(* IEC 61131-3 sources: NachHouse_TST/OSCAT_BasicLib/OscatBasicLib_333a (part 5) *)

(* ---- Plc_Time.ST ---- *)
(* @PATH := '\/Engineering\/measurements' *)
FUNCTION T_PLC_MS : DWORD
(*
  T_PLC_MS reads the internal PLC timer and return the time, it has the advantage to be able to set a debug mode
  and speed up the counter to test the plc timer overrun which occurs every 50 days respectively 25 days at siemens S7
  this routine also allows to correct the behavior of s7 where the internal plc counter will not count all 32 bits.

  version 1.2 16. nov 2008
  programmer  hugo
  tested by oscat
*)
  VAR CONSTANT
    debug : BOOL := 0;
    N : INT := 0;
    offset : DWORD := 0;
  END_VAR
  VAR
  //  tx : TIME;
  END_VAR
  VAR_EXTERNAL
    AT %SL52 : DWORD;
  END_VAR
  VAR_TEMP
    temp : DWORD;
  END_VAR

  //???tx := TIME();
  T_PLC_MS := %SL52;
  (* hier muss die korrektur für step7 stattfinden
  plctime muss den vollen wertebereich von time ausnutzen:
  wenn bei step7 time -24tage bis plus 24 tage ist dann muss der timer auch beim überlauf auf -24tage springen
  und auf keinen fall auf 0 !!!!
  für siemens muss ein weiterer fb im main eingebunden werden der sicherstellt das alle 32 bits durchgezählt werden.
  es kann nur ein fb sein den er muss sich das oberste (32te) bit merken.
  oder etwa spring s7 bei überlauf auf -24 tage????? dann wäre keine korrektur nötig.
  *)
  IF debug THEN
    //???  T_PLC_MS := (SHL(T_PLC_MS,N) OR SHL(DWORD#1,N)-1) + OFFSET;
    temp := UDINT_TO_DWORD( DWORD_TO_UDINT( SHL(DWORD#1,INT_TO_UINT(N))) -1);
    temp := temp OR SHL(%SL52,INT_TO_UINT(N));
    T_PLC_MS := UDINT_TO_DWORD( DWORD_TO_UDINT(temp) + DWORD_TO_UDINT(OFFSET));
  END_IF;

(* revision history
  hm  14.9.2007 rev 1.0
    original version

  hm  12. nov 2007  rev 1.1
    added temporaray variable tx because some compilers could not handle time() as an argument

  hm  16. nov. 2008 rev 1.2
    initialized constants with 0 for compatibility reasons
*)
END_FUNCTION

(* @PATH := '\/Engineering\/measurements' *)
FUNCTION T_PLC_US : DWORD
(*
  T_PLC_US reads the internal PLC timer and return the time, it has the advantage to be able to set a debug mode
  and speed up the counter to test the plc timer overrun which occurs every 50 days respectively 25 days at siemens S7
  this routine also allows to correct the behavior of s7 where the internal plc counter will not count all 32 bits.

  version 1.2 16 nov 2008
  programmer  hugo
  tested by tobias
*)
  VAR CONSTANT
    debug : BOOL := 0;
    N : INT := 0;
    offset : DWORD := 0;
  END_VAR
  VAR
  //  tx : TIME;
  END_VAR
  VAR_EXTERNAL
    AT %SL52 : DWORD;
  END_VAR
  VAR_TEMP
    temp : DWORD;
    temp_T_PLC_US : DWORD;
  END_VAR

  //???tx := TIME();
  //???T_PLC_US := TIME_TO_DWORD(Tx)*1000;
  T_PLC_US := UDINT_TO_DWORD(DWORD_TO_UDINT(%SL52)*1000);
  (* hier muss die korrektur für step7 stattfinden
  plctime muss den vollen wertebereich von time ausnutzen:
  wenn bei step7 time -24tage bis plus 24 tage ist dann muss der timer auch beim überlauf auf -24tage springen
  und auf keinen fall auf 0 !!!!
  für siemens muss ein weiterer fb im main eingebunden werden der sicherstellt das alle 32 bits durchgezählt werden.
  es kann nur ein fb sein den er muss sich das oberste (32te) bit merken.
  oder etwa spring s7 bei überlauf auf -24 tage????? dann wäre keine korrektur nötig.
  *)
  IF debug THEN
    //???T_PLC_US := (SHL(T_PLC_US,N) OR SHL(DWORD#1,N)-1) + OFFSET;
    temp_T_PLC_US := UDINT_TO_DWORD(DWORD_TO_UDINT(%SL52)*1000);
    temp := UDINT_TO_DWORD( DWORD_TO_UDINT( SHL(DWORD#1,INT_TO_UINT(N))) -1);
    temp := temp OR SHL(temp_T_PLC_US,INT_TO_UINT(N));
    T_PLC_US := UDINT_TO_DWORD( DWORD_TO_UDINT(temp) + DWORD_TO_UDINT(OFFSET));
  END_IF;

(* revision history
  hm  14.9.2007 rev 1.0
    original version

  hm  12. nov 2007  rev 1.1
    added temporaray variable tx because some compilers could not handle time() as an argument

  hm  16. nov. 2008 rev 1.2
    initialized constants with 0 for compatibility reasons
*)
END_FUNCTION

(* @PATH := '\/String' *)
FUNCTION TO_UPPER : BYTE
(*
  to_upper converts a character from lowercase to uppercase

  version 1.3 16. jan. 2009
  programmer  hugo
  tested by   oscat
*)
  VAR_INPUT
    IN : BYTE;
  END_VAR

  IF (in > 96) AND (in < 123) THEN
     TO_UPPER := in AND 16#DF;
  ELSIF (in > 223) AND (in <> 247) AND (in <> 255) AND setup.EXTENDED_ASCII THEN
     TO_UPPER := in AND 16#DF;
  ELSE
     TO_UPPER := in;
  END_IF;

(* revision history
  hm  6. mar. 2008  rev 1.0
    original version

  hm  19. oct. 2008 rev 1.1
    changed setup constants

  ks  25. oct. 2008 rev 1.2
    optimized code

  hm 16. jan 2009 rev 1.3
    corrected an error in module
  *)
END_FUNCTION

(* ---- Sensors.ST ---- *)
(* @PATH := '\/Engineering\/sensor' *)
FUNCTION MULTI_IN : REAL
(*
  multi_in is a signal conditioning function which can be configured in 8 different ways.
  it is used to read multiple sensors for the same value and protect the user from broken sensors or invalid data from sensors.

  multi_in can be configured in different ways:
    mode = 0 means the the avg of the 3 inputs is used, this mode is the default mode.
    mode = 1 means in_1 is used.
    mode = 2 means in_2 is used.
    mode = 3 means in_3 is used.
    mode = 4 means default is used.
    mode = 5 means the lowest of the 3 external temperatures is used.
    mode = 6 means the higest externnal temperature is used.
    mode = 7 means the midlle input is used, if there are only two working, the lowest input is used.
    mode > 7 ,eans output is 0 at all times.
    in any config mode, an input higher then in_max or lower then in_min is ignored to prevent values from broken sensors or wires.
    if all inputs are higher then in_max or lower then in_min, a default value (default) is used.

  version 1.4 18. jul. 2009
  programmer  oscat
  tested by   oscat
*)
  VAR_INPUT
    in_1 : REAL;
    in_2 : REAL;
    in_3 : REAL;
    default : REAL;
    in_min : REAL;
    in_max : REAL;
    mode : BYTE;
  END_VAR
  VAR
    count: INT;
    F1: BOOL;
    F2: BOOL;
    F3: BOOL;
  END_VAR

  F1 :=  in_1 > in_min AND in_1 < in_max;
  F2 :=  in_2 > in_min AND in_2 < in_max;
  F3 :=  in_3 > in_min AND in_3 < in_max;

  CASE BYTE_TO_USINT(mode) OF
  0:  count := 0;
    IF F1 THEN
      count := count + 1;
      MULTI_IN := in_1;
    ELSE
      MULTI_IN := 0.0;
    END_IF;
    IF F2 THEN
      count := count + 1;
      MULTI_IN := MULTI_IN + in_2;
    END_IF;
    IF F3 THEN
      count := count + 1;
      MULTI_IN := MULTI_IN + in_3;
    END_IF;
    MULTI_IN := SEL(count = 0, MULTI_IN / INT_TO_REAL(count), default);

  1:  MULTI_IN := SEL(F1, default, IN_1);

  2:  MULTI_IN := SEL(F2, default, IN_2);

  3:  MULTI_IN := SEL(F3, default, IN_3);

  4:  MULTI_IN := default;

  5:  MULTI_IN := SEL(F1, in_max, IN_1);
    IF F2 AND in_2 < MULTI_IN THEN MULTI_IN := in_2; END_IF;
    IF F3 AND in_3 < MULTI_IN THEN MULTI_IN := in_3; END_IF;
    IF MULTI_IN = in_max THEN MULTI_IN := default; END_IF;

  6:  MULTI_IN := SEL(F1, in_min, IN_1);
    IF F2 AND in_2 > MULTI_IN THEN MULTI_IN := in_2; END_IF;
    IF F3 AND in_3 > MULTI_IN THEN MULTI_IN := in_3; END_IF;
    IF MULTI_IN = in_min THEN MULTI_IN := default; END_IF;

  7:  IF F1 AND F2 AND F3 THEN MULTI_IN := MID3(in_1, in_2, in_3);
    ELSIF F1 AND F2 THEN MULTI_IN := MIN(in_1, in_2);
    ELSIF F1 AND F3 THEN MULTI_IN := MIN(in_1, in_3);
    ELSIF F2 AND F3 THEN MULTI_IN := MIN(in_2, in_3);
    ELSIF F1 THEN MULTI_IN := in_1;
    ELSIF F2 THEN MULTI_IN := in_2;
    ELSIF F3 THEN MULTI_IN := in_3;
    ELSE MULTI_IN := default;
    END_IF;
  ELSE
    MULTI_IN := 0.0;
  END_CASE;

(*
  hm 1.1.2007   rev 1.1
    changed midr to mid3 function

  hm  14. 10. 2008  rev 1.2
    corrected an error for in_3 overrange detection
    improved performance

  hm  11. mar. 2009 rev 1.3
    changed real constants to use dot syntax

  hm  18. jul. 2009 rev 1.4
    improved performance
*)
END_FUNCTION

(* @PATH := '\/Engineering\/sensor' *)
FUNCTION RES_NI : REAL
(*
  this function returs the resistance for a nickel sensor for a temperature range from -60..+180 °C

  version 1.2 2 dec 2007
  programmer  hugo
  tested by   tobias
*)
  VAR_INPUT
    T : REAL;
    R0 : REAL;
  END_VAR
  VAR CONSTANT
    A : REAL := 0.5485;
    B : REAL := 0.665E-3;
    C : REAL := 2.805E-9;
  END_VAR
  VAR
    T2: REAL;
  END_VAR

  T2 := T * T;
  RES_NI := R0 + A * T + B * T2 + C * T2 * T2;

(* revision history
  hm  4.8.2006    rev 1.0
    original version

  hm  13.9.2007   rev 1.1
    changed coding for better performance

  hm  2. dec. 2007  rev 1.2
    changed code for better performance
*)
(*
 Auszug aus DIN 43760 für Ni100

°C    R   °C    R   °C  R   °C    R   °C    R

-60   69,5  -10   94,6  40  123,0   90    154,9   140   190,9
-55   71,9  -5    97,3  45  126,0   95    158,3   145   194,8
-50   74,3  0     100,0   50  129,1   100   161,8   150   198,7
-45   76,7  5     102,8   55  132,2   105   165,3   155   202,6
-40   79,1  10    105,6   60  135,3   110   168,8   160   206,6
-35   81,6  15    108,4   65  138,5   115   172,4   165   210,7
-30   84,2  20    111,2   70  141,7   120   176,0   170   214,8
-25   86,7  25    114,1   75  145,0   125   179,6   175   219,0
-20   89,3  30    117,1   80  148,3   130   183,3   180   223,2
-15   91,9  35    120,0   85  151,6   135   187,1
*)
END_FUNCTION

(* @PATH := '\/Engineering\/sensor' *)
FUNCTION RES_NTC : REAL
(*
  this function returs the resistance for a NTC sensor for a given temperature in °C.
  RN is the resistance at 25 °C and B is a constant for the given sensor.

  version 1.1 11. mar. 2009
  programmer  hugo
  tested by   tobias
*)
  VAR_INPUT
    T : REAL;
    RN : REAL;
    B : REAL;
  END_VAR

  RES_NTC := RN * EXP(B * (1.0 / (T+273.15) - 0.00335401643468053));

(* revision history
  hm 30. dec. 2008  rev 1.0
    original version

  hm  11. mar. 2009 rev 1.1
    changed real constants to use dot syntax
*)
END_FUNCTION

(* @PATH := '\/Engineering\/sensor' *)
FUNCTION RES_PT : REAL
(*
  this function returs the resistance for a platinum sensor for a temperature range from -200..+850 °C

  version 1.3 11. mar. 2009
  programmer  hugo
  tested by   oscat
*)
  VAR_INPUT
    T : REAL;
    R0 : REAL;
  END_VAR
  VAR CONSTANT
    A : REAL := 3.90802E-3 ;
    B : REAL := -5.802E-7;
    C : REAL := -4.27350E-12;
  END_VAR
  VAR
    T2: REAL;
  END_VAR

  T2 := T * T;

  IF T >= 0.0 THEN
    RES_PT := R0 * ( 1.0 + A * T + B * T2);
  ELSE
    RES_PT := R0 * ( 1.0 + A * T + B * T2 + C * (T - 100.0) * T2 * T);
  END_IF;

(* revision history
  hm  4. aug. 2006  rev 1.1
    original version

  hm  2. dec 2007 rev 1.2
    changed code for better performance

  hm  11. mar. 2009 rev 1.3
    changed real constants to use dot syntax
*)
(*
 Auszug aus DIN 43760 für Pt100

°C    R   °C    R   °C  R     °C    R     °C    R     °C    R

-200  18,49   -100  60,25   0   100,00  100   138,50  200   175,84  300   212,02
-195  20,65   -95   62,28   5   101,95  105   140,39  205   177,68  305   213,80
-190  22,80   -90   64,30   10  103,90  110   142,29  210   179,51  310   215,57
-185  24,94   -85   66,31   15  105,85  115   144,17  215   181,34  315   217,35
-180  27,08   -80   68,33   20  107,79  120   146,06  220   183,17  320   219,12
-175  29,20   -75   70,33   25  109,73  125   147,94  225   184,99  325   220,88
-170  31,32   -70   72,33   30  111,67  130   149,82  230   186,82  330   222,65
-165  33,43   -65   74,33   35  113,61  135   151,70  235   188,63  335   224,41
-160  35,33   -60   76,33   40  115,54  140   153,58  240   190,45  340   226,17
-155  37,63   -55   78,32   45  117,47  145   155,45  245   192,26  345   227,92
-150  39,71   -50   80,31   50  119,40  150   157,31  250   194,07  350   229,67
-145  41,79   -45   82,29   55  121,32  155   159,18  255   195,88  355   231,42
-140  43,87   -40   84,27   60  123,24  160   161,04  260   197,69  360   233,17
-135  45,94   -35   86,25   65  125,16  165   162,90  265   199,49  365   234,91
-130  48,00   -30   88,22   70  127,07  170   164,76  270   201,29  370   236,65
-125  50,06   -25   90,19   75  128,98  175   166,61  275   203,08  375   238,39
-120  52,11   -20   92,16   80  130,89  180   168,46  280   204,88  380   240,13
-115  54,15   -15   94,12   85  132,80  185   170,31  285   206,67  385   241,86
-110  56,19   -10   96,09   90  134,70  190   172,16  290   208,45  390   243,59
-105  58,22   -5    98,04   95  136,60  195   174,00  295   210,24  395   245,31
*)
END_FUNCTION

(* @PATH := '\/Engineering\/sensor' *)
FUNCTION RES_SI : REAL
(*
  this function returs the resistance for a silicon sensor for a temperature range from -50..+150 °C
  for example KTY10 normaly Rs at 25 °C

  version 1.2 11. mar. 2009
  programmer  hugo
  tested by   tobias
*)
  VAR_INPUT
    T : REAL;
    RS : REAL;
    TS : REAL;
  END_VAR
  VAR CONSTANT
    A : REAL := 7.64E-3;
    B : REAL := 1.66E-5;
  END_VAR
  VAR
    TX: REAL;
  END_VAR

  TX := T - TS;
  RES_SI := RS * ( 1.0 + A * TX + B * TX * TX);

(* revision history
  hm  4. aug 2006 rev 1.0
    original version

  hm  2. dec 2007 rev 1.1
    changed code for better performance

  hm  11. mar. 2009 rev 1.2
    changed real constants to use dot syntax
*)
END_FUNCTION

(* @PATH := '\/Engineering\/sensor' *)
FUNCTION SENSOR_INT : REAL
(*
  this function calculates the real resistance of a sensor RX given a parasitic resistor in parallel to the sensor and an additional serial resistor.
  for example a parasitic parallel resistor for a PT100 can be ignored but a series resistor is the cable to the sensor.
  for a humidity sensor, the parallel resistor is more dramatic and needs to be considered.
  the function allows to consider a parallel and serial resistor at the same time.
  with this function and known parasitic serial and parallel resistors the true resistance of the sensor can be calculated.

  version 1.3 11. mar. 2009
  programmer  hugo
  tested by   tobias
*)
  VAR_INPUT
    Voltage : REAL;
    Current : REAL;
    RP : REAL;
    RS : REAL;
  END_VAR
  VAR
    RG: REAL;
  END_VAR

  IF current <> 0.0 THEN
    RG := voltage / current;
    SENSOR_INT := RP * ( RG - RS) / ( RP + RS - RG);
  END_IF;

(* revisaion history
  hm 20.1.2007    rev 1.1
    deleted input R0 which was not needed.

  hm  2. dec 2007 rev 1.2
    corrected an error in formula and improoved speed

  hm  11. mar. 2009 rev 1.3
    changed real constants to use dot syntax
*)
END_FUNCTION

(* @PATH := '\/Engineering\/sensor' *)
FUNCTION TEMP_NI : REAL
(*
  this function returns the temperature for a nickel sensor in a range from -60..+180 °C

  version 1.5 10. mar. 2009
  programmer  hugo
  tested by   tobias
*)
  VAR_INPUT
    Res : REAL;
    R0 : REAL;
  END_VAR

  TEMP_NI := (SQRT(0.30085225 - 2.66E-3 * (R0 - Res)) - 0.5485) * 751.8796992;

(* revision history
  hm 24.1.2007    rev 1.1
    deleted unused variable A, B, C

  hm 10.9.2007    rev 1.2
    changed accuracy to 0.02 degrees to improove performace

  hm 17. 12 2007  rev 1.3
    improovements for better performance and higher accuracy

  hm  6. jan 2008 rev 1.4
    further performance improvement

  hm  10. mar. 2009 rev 1.5
    removed nested comments
*)
END_FUNCTION

(* @PATH := '\/Engineering\/sensor' *)
FUNCTION TEMP_NTC : REAL
(*
  this function returs the temperature for a NTC sensor for a range from 0..85 °C.
  RN is the resistance at 25 °C and B is a constant for the given sensor.

  version 1.1 11. mar. 2009
  programmer  hugo
  tested by   tobias
*)
  VAR_INPUT
    RES : REAL;
    RN : REAL;
    B : REAL;
  END_VAR

  IF res > 0.0 THEN
    TEMP_NTC := B * 298.15 / (B + LN(RES / RN) * 298.15) -273.15;
  END_IF;

(* revision history
  hm 30. dec. 2008  rev 1.0
    original version

  hm  11. mar. 2009 rev 1.1
    changed real constants to use dot syntax
*)
END_FUNCTION

(* @PATH := '\/Engineering\/sensor' *)
FUNCTION TEMP_PT : REAL
(*
  this function returs the temperature for a platinum sensor for a range from -200..+850 °C

  version 1.7 11. mar. 2009
  programmer  hugo
  tested by   oscat
*)
  VAR_INPUT
    Res : REAL;
    R0 : REAL;
  END_VAR
  VAR CONSTANT
    A : REAL := 3.9083E-3 ;
    B : REAL := -5.775E-7;
    accuracy : REAL := 0.01;
  END_VAR
  VAR
    step: REAL := 50.0;
    X: REAL;
    Y: REAL;
    t1: REAL;
    pt : PTR_TO UDINT; //DWORD;
  END_VAR
  VAR_TEMP
    tmp : REAL;
  END_VAR

  X := A * R0;
  Y := B * R0;
  IF Res >= R0 THEN
    t1 := X * X - 4.0 * Y * (R0 - Res);
    IF t1 < 0.0 THEN
      tmp := 10000.0;
    ELSE
      tmp := (-X + SQRT(t1)) / (2.0 * Y);
    END_IF;
  ELSE
    pt := ADR(step);
    (* since the formula cannot be solved this is a successive approximation *)
    tmp := -100.0;
    WHILE step > accuracy DO
      (* test if result greater or less *)
      IF RES_PT(tmp, R0) < res THEN tmp := tmp + step; ELSE tmp := tmp - step; END_IF;
      pt^ := pt^ - 8388608;  (* this is a super fast divide by 2 method for non floating point CPUs *)
      (* the alternative code: step := step * 0.5; *)
    END_WHILE;
  END_IF;
  TEMP_PT := tmp;

(* revision history
  rev 1.1 hm 24.1.2007
    deleted unused variable C

  rev 1.2 hm 10.9.2007
    reduced accuracy to 0.02 to shorten execution time

  rev 1.3 hm  2. dec 2007
    changed code for better performance

  rev 1.4 hm  23. dec 2007
    avoid a negative square root if input values are wrong

  rev 1.5 hm  5. jan 2008
    replaced / 2 with * 0.5 for better performance

  hm  31. oct. 2008 rev 1.6
    improved performance

  hm  11. mar. 2009 rev 1.7
    changed real constants to use dot syntax
*)
END_FUNCTION

(* @PATH := '\/Engineering\/sensor' *)
FUNCTION TEMP_SI : REAL
(*
  this function returs the temperature for a silicon sensor for a range from -60..+180 °C
  for example KTY10 RS at TS normally 25 °C

  version 1.5 10. mar. 2009
  programmer  hugo
  tested by   tobias
*)
  VAR_INPUT
    Res : REAL;
    RS : REAL;
    TS : REAL;
  END_VAR

  TEMP_SI := (-7.64E-3 + SQRT(Res / RS * 6.64E-5 - 0.803E-5)) * 30120.48193 + TS;

(* revision history
  hm 24.1.2007    rev 1.1
    the function would only work for TS = 25, now it works for other values of ts.

  hm 10.9.2007    rev 1.2
    changed the function to use successive approcimation to avoid an error generated by a sqrt from a negative result.
    changed accuracy to 0.02 degrees to shorten execution time

  hm 17. 12 2007  rev 1.3
    improovements for better performance

  hm  6. jan 2008 rev 1.4
    further performance improvement

  hm  10. mar. 2009 rev 1.5
    removed nested comments
*)
END_FUNCTION

(* ---- String.ST ---- *)
(* @NESTEDCOMMENTS := 'Yes' *)
(* @PATH := '\/String' *)
(* @OBJECTFLAGS := '0, 8' *)
(* @SYMFILEFLAGS := '2048' *)
FUNCTION TO_UPPER : BYTE
(*
  to_upper converts a character from lowercase to uppercase

  version 1.3 16. jan. 2009
  programmer  hugo
  tested by   oscat
*)
  VAR_INPUT
    IN : BYTE;
  END_VAR

  (* @END_DECLARATION := '0' *)
  IF BYTE_TO_USINT(in) > 96 AND BYTE_TO_USINT(in) < 123 THEN
     TO_UPPER := in AND 16#DF;
  ELSIF BYTE_TO_USINT(in) > 223 AND BYTE_TO_USINT(in) <> 247 AND BYTE_TO_USINT(in) <> 255 AND setup.EXTENDED_ASCII THEN
     TO_UPPER := in AND 16#DF;
  ELSE
     TO_UPPER := in;
  END_IF;

  (* revision history
  hm  6. mar. 2008  rev 1.0
    original version

  hm  19. oct. 2008 rev 1.1
    changed setup constants

  ks  25. oct. 2008 rev 1.2
    optimized code

  hm 16. jan 2009 rev 1.3
    corrected an error in module

  *)
END_FUNCTION

(* ---- Vector_Mathematics.ST ---- *)
(* @PATH := '\/Mathematical\/Vektormathematik' *)
FUNCTION V3_ABS : REAL
(*
  this function calculates the length of a vectors in a 3 dimensional space

  version 1.0 11 dec 2007
  programmer  hugo
  tested by   tobias
*)
  VAR_INPUT
    A : Vector_3;
  END_VAR

  V3_ABS := SQRT(A.X * A.X + A.Y * A.Y + A.Z * A.Z);

(* revision history
  hm  11 dec 2007 rev 1.0
      original version
*)
END_FUNCTION

(* @PATH := '\/Mathematical\/Vektormathematik' *)
FUNCTION V3_ADD : vector_3
(*
  this function adds two vectors in a 3 dimensional space

  version 1.0 11 dec 2007
  programmer  hugo
  tested by   tobias
*)
  VAR_INPUT
    A : Vector_3;
    B : Vector_3;
  END_VAR

  V3_ADD.X := A.X + B.X;
  V3_ADD.Y := A.Y + B.Y;
  V3_ADD.Z := A.Z + B.Z;

(* revision history
  hm    11 dec 2007 rev 1.0
        original version
*)
END_FUNCTION

(* @PATH := '\/Mathematical\/Vektormathematik' *)
FUNCTION V3_DPRO : REAL
(*
  this function calculates the dot product of two vectors in 3 dimensional space

  version 1.0 11 dec 2007
  programmer  hugo
  tested by   tobias
*)
  VAR_INPUT
    A : Vector_3;
    B : Vector_3;
  END_VAR

  V3_DPRO := A.X * B.X + A.Y * B.Y + A.Z * B.Z;

(* revision history
  hm  11 dec 2007 rev 1.0
      original version
*)
END_FUNCTION

(* @PATH := '\/Mathematical\/Vektormathematik' *)
FUNCTION V3_ANG : REAL
(*
  this function calculates the angle between two vectors in a 3 dimensional space

  version 1.1 10. mar. 2009
  programmer  hugo
  tested by   tobias
*)
  VAR_INPUT
    A : Vector_3;
    B : Vector_3;
  END_VAR
  VAR
    d : REAL;
  END_VAR

  d := V3_ABS(A) * V3_ABS(B);
  IF d > 0.0 THEN
    V3_ANG := ACOS(LIMIT(-1.0, V3_DPRO(A, B) / d,1.0));
  END_IF;

(* revision history
  hm  11. dec. 2007 rev 1.0
    original version

  hm  10. mar. 2009 rev 1.1
    changed syntax of real constants to 0.0
*)
END_FUNCTION

(* @PATH := '\/Mathematical\/Vektormathematik' *)
FUNCTION V3_SMUL : vector_3
(*
  this function multiplies a vectors in a 3 dimensional space with a skalar M

  version 1.0 11 dec 2007
  programmer  hugo
  tested by   tobias
*)
  VAR_INPUT
    A : Vector_3;
    M : REAL;
  END_VAR

  V3_SMUL.X := A.X * M;
  V3_SMUL.Y := A.Y * M;
  V3_SMUL.Z := A.Z * M;

(* revision history
  hm    11 dec 2007 rev 1.0
        original version
*)
END_FUNCTION

(* @PATH := '\/Mathematical\/Vektormathematik' *)
FUNCTION V3_NORM : vector_3
(*
  this function generates a vectors with absolute length 1 from a vector A in a 3 dimensional space

  version 1.1 10. mar. 2009
  programmer  hugo
  tested by   tobias
*)
  VAR_INPUT
    A : Vector_3;
  END_VAR
  VAR
    la: REAL;
  END_VAR

  la := V3_ABS(A);
  IF la > 0.0 THEN
    V3_NORM := V3_SMUL(A, 1.0 / la);
  END_IF;

(* revision history
  hm  11 dec 2007 rev 1.0
    original version

  hm  10. mar. 2009 rev 1.1
    changed syntax of real constants to 0.0
*)
END_FUNCTION

(* @PATH := '\/Mathematical\/Vektormathematik' *)
FUNCTION V3_NUL : BOOL
(*
  this function checks if a vectors in a null Vector

  version 1.1 10. mar. 2009
  programmer  hugo
  tested by   tobias
*)
  VAR_INPUT
    A : Vector_3;
  END_VAR

  V3_NUL := A.X = 0.0 AND A.Y = 0.0 AND A.Z = 0.0;

(* revision history
  hm  12 dec 2007 rev 1.0
    original version

  hm  10. mar. 2009 rev 1.1
    changed syntax of real constants to 0.0
*)
END_FUNCTION

(* @PATH := '\/Mathematical\/Vektormathematik' *)
FUNCTION V3_XPRO : vector_3
(*
  this function adds two vectors in a 3 dimensional space

  version 1.0 11 dec 2007
  programmer  hugo
  tested by   tobias
*)
  VAR_INPUT
    A : Vector_3;
    B : Vector_3;
  END_VAR

  V3_XPRO.X := A.Y * B.Z - A.Z * B.Y;
  V3_XPRO.Y := A.Z * B.X - A.X * B.Z;
  V3_XPRO.Z := A.X * B.Y - A.Y * B.X;

(* revision history
  hm    11 dec 2007 rev 1.0
    original version
*)
END_FUNCTION

(* @PATH := '\/Mathematical\/Vektormathematik' *)
FUNCTION V3_PAR : BOOL
(*
  this function checks if two vectors in a 3 dimensional space are parallel.
  which means the two vectors have the same direction

  version 1.1 10. mar. 2009
  programmer  hugo
  tested by   tobias
*)
  VAR_INPUT
    A : Vector_3;
    B : Vector_3;
  END_VAR

  V3_PAR := V3_ABS(V3_XPRO(A, B)) = 0.0;

(* revision history
  hm  11 dec 2007 rev 1.0
    original version

  hm  10. mar. 2009 rev 1.1
    changed syntax of real constants to 0.0
*)
END_FUNCTION

(* @PATH := '\/Mathematical\/Vektormathematik' *)
FUNCTION V3_REV : vector_3
(*
  this function reverses a vector in a 3 dimensional space

  version 1.0 11 dec 2007
  programmer  hugo
  tested by   tobias
*)
  VAR_INPUT
    A : Vector_3;
  END_VAR

  V3_REV.X := -A.X;
  V3_REV.Y := -A.Y;
  V3_REV.Z := -A.Z;

(* revision history
  hm    11 dec 2007 rev 1.0
        original version
*)
END_FUNCTION

(* @PATH := '\/Mathematical\/Vektormathematik' *)
FUNCTION V3_SUB : vector_3
(*
  this function subtracts two vectors in a 3 dimensional space
  V3_SUB = A - B

  version 1.0 11 dec 2007
  programmer  hugo
  tested by   tobias
*)
  VAR_INPUT
    A : Vector_3;
    B : Vector_3;
  END_VAR

  V3_SUB.X := A.X - B.X;
  V3_SUB.Y := A.Y - B.Y;
  V3_SUB.Z := A.Z - B.Z;

(* revision history
  hm    11 dec 2007 rev 1.0
    original version
*)
END_FUNCTION

(* @PATH := '\/Mathematical\/Vektormathematik' *)
FUNCTION V3_XANG : REAL
(*
  this function calculates the angle between the X-axis and a vectors in a 3 dimensional space

  version 1.1 10. mar. 2009
  programmer  hugo
  tested by   tobias
*)
  VAR_INPUT
    A : Vector_3;
  END_VAR
  VAR
    la: REAL;
  END_VAR

  la := V3_ABS(a);
  IF la > 0.0 THEN
    V3_XANG := ACOS(A.X / la);
  END_IF;

(* revision history
  hm  11 dec 2007 rev 1.0
    original version

  hm  10. mar. 2009 rev 1.1
    changed syntax of real constants to 0.0
*)
END_FUNCTION

(* @PATH := '\/Mathematical\/Vektormathematik' *)
FUNCTION V3_YANG : REAL
(*
  this function calculates the angle between the Y-axis and a vectors in a 3 dimensional space

  version 1.1 10. mar. 2009
  programmer  hugo
  tested by   tobias
*)
  VAR_INPUT
    A : Vector_3;
  END_VAR
  VAR
    la: REAL;
  END_VAR

  la := V3_ABS(a);
  IF la > 0.0 THEN
    V3_YANG := ACOS(A.Y / la);
  END_IF;

(* revision history
  hm  11 dec 2007 rev 1.0
    original version

  hm  10. mar. 2009 rev 1.1
    changed syntax of real constants to 0.0
*)
END_FUNCTION

(* @PATH := '\/Mathematical\/Vektormathematik' *)
FUNCTION V3_ZANG : REAL
(*
  this function calculates the angle between the Z-axis and a vectors in a 3 dimensional space

  version 1.1 10. mar. 2009
  programmer  hugo
  tested by   tobias
*)
  VAR_INPUT
    A : Vector_3;
  END_VAR
  VAR
    la: REAL;
  END_VAR

  la := V3_ABS(a);
  IF la > 0.0 THEN
    V3_ZANG := ACOS(A.Z / la);
  END_IF;

(* revision history
  hm  11 dec 2007 rev 1.0
    original version

  hm  10. mar. 2009 rev 1.1
    changed syntax of real constants to 0.0
*)
END_FUNCTION

(* ---- Arithmetic_Functions.ST ---- *)
TYPE
  OSCAT_BASIC_ARRAY1_20x0_1_OF_REAL : ARRAY[1..20, 0..1] OF REAL;
END_TYPE

(* @PATH := '\/Mathematical\/functions' *)
FUNCTION F_LIN : REAL
(*
  this function calculates the linear equation f_lin = a*x + b

  version 1.0 1 sep 2006
  programmer  hugo
  tested by   tobias
*)
  VAR_INPUT
    X : REAL;
    A : REAL;
    B : REAL;
  END_VAR

  F_lin := A * X + B;
END_FUNCTION

(* @PATH := '\/Mathematical\/functions' *)
FUNCTION F_LIN2 : REAL
(*
  this function calculates the linear equation f_lin = a*x + b given by two points x1/y1 and x2/y2.

  version 1.0 1 jan 2007
  programmer  hugo
  tested by   tobias
*)
  VAR_INPUT
    X : REAL;
    X1: REAL;
    Y1 : REAL;
    X2 : REAL;
    Y2 : REAL;
  END_VAR

  F_LIN2 := (Y2 - Y1) / (X2 - X1) * (X - X1) + Y1;

(* revision history
  hm  1. jan. 2007  rev 1.0
    original release

  hm  17. dec. 2008 rev 1.1
    optimized formula
*)
END_FUNCTION

(* @PATH := '\/Mathematical\/functions' *)
FUNCTION F_POLY : REAL
(*
  this function calculates the polynom C[0] + C[1]*X^1 + C[2]*X^2 * C[3]*X^3 + C[4]*X^4 + C[5]*X^5 + C[6]*X^6 + C[7]*X^7

  version 1.1 18. mar. 2011
  programmer  hugo
  tested by   tobias
*)
  VAR_INPUT
    X : REAL;
    C : ARRAY[0..7] OF REAL;
  END_VAR

  F_POLY := ((((((( c[7] * x + c[6] ) * x + c[5] ) * x + c[4] ) * x + c[3] ) * x + c[2] ) * x + c[1] ) * x + c[0] ) ;

(* revision history
  hm    20. may. 2008   rev 1.0
    original version

  hm  18. mar. 2011 rev 1.1
    improved performance
*)
END_FUNCTION

(* @PATH := '\/Mathematical\/functions' *)
FUNCTION F_POWER : REAL
(*
  this function calculates the power equation f_power = a*x^n

  version 1.0 1 sep 2006
  programmer  hugo
  tested by   tobias
*)
  VAR_INPUT
    a : REAL;
    x : REAL;
    n : REAL;
  END_VAR

  F_POWER := a * EXPT(X, N);
END_FUNCTION

(* @PATH := '\/Mathematical\/functions' *)
FUNCTION F_QUAD : REAL
(*
  this function calculates the quadratic equation f_lin = a*x + b

  version 1.1 18. Mar. 2011
  programmer  hugo
  tested by   tobias
*)
  VAR_INPUT
    X : REAL;
    A : REAL;
    B : REAL;
    C : REAL;
  END_VAR

  F_QUAD :=  (A * X + B) * X + C;

(* revision history
  hm  1. sep. 2006  rev 1.0
    original version

  hm  18. mar. 2001 rev 1.1
    improved performance
*)
END_FUNCTION

(* @PATH := '\/Mathematical\/functions' *)
FUNCTION FRMP_B : BYTE
(*
  this function calculates a ramp and limits the output to 0 .. 255 without overflow problems

  version 1.0   17. feb. 2011
  programmer  hugo
  tested by   oscat
*)
  VAR_INPUT
    START : BYTE;
    DIR : BOOL;
    TD : TIME;
    TR : TIME;
  END_VAR
  VAR
    tmpw : DWORD;
    tmpb : BYTE;
  END_VAR

  IF TD < TR THEN
    //???FRMP_B := MIN(DWORD_TO_BYTE(SHL(TIME_TO_DWORD(TD), 8) / TIME_TO_DWORD(TR)), SEL(DIR, START, BYTE#255 - START));
    tmpw := SHL(TIME_TO_DWORD(TD), 8);
    tmpw := UDINT_TO_DWORD( DWORD_TO_UDINT(tmpw) /  TIME_TO_UDINT(TR));
    tmpb := MIN( DWORD_TO_BYTE(tmpw), SEL( DIR, START, USINT_TO_BYTE(USINT#255 - BYTE_TO_USINT(START))));
    IF DIR THEN
      FRMP_B := USINT_TO_BYTE( BYTE_TO_USINT(START) + BYTE_TO_USINT(tmpb));
    ELSE
      FRMP_B := USINT_TO_BYTE( BYTE_TO_USINT(START) - BYTE_TO_USINT(tmpb));
    END_IF;
  ELSE
    FRMP_B := SEL(DIR, 0, 255);
  END_IF;

(* revision history
  17. feb. 2011 rev 1.0
    new module
*)
END_FUNCTION

(* @PATH := '\/Mathematical\/functions' *)
FUNCTION_BLOCK FT_AVG
(*
  this function calculates the moving average over n samples from a sequential input
  the input values are shifted into an N deep buffer and the avg of this buffer is diplayed at anytime on the output.
  a rst will load the buffer with the current in value..

  version 1.5 10. mar. 2009
  programmer  hugo
  tested by   oscat
*)
  VAR_INPUT
    IN : REAL;
    E : BOOL := TRUE;
    N : INT := 32;
    RST : BOOL;
  END_VAR
  VAR_OUTPUT
    AVG : REAL;
  END_VAR
  VAR
    buff : DELAY;
    i: INT;
    init : BOOL;
  END_VAR

  (* limit n to a max of 32 because delay can do max 32 cycles *)
  buff.N := LIMIT(0, N, 32);

  IF NOT init OR rst THEN
    FOR i := 1 TO N DO
      buff(in := in);
    END_FOR;
    avg := in;
    init := TRUE;
  ELSIF E THEN
    buff(in := in);
    avg := avg + (in - buff.out ) / INT_TO_REAL(N);
  END_IF;

(* revision history
  hm  7. jan. 2007  rev 1.1
    chaged rst logic to load the buffer with the actual input value instead of 0.
    added en input to allow better control of signal flow
    added init to load the buffer with in at startup to avoid rampup at beginning.
    deleted unused variable cnt.

  hm  14. jun. 2008 rev 1.2
    set default for input en = TRUE and N = 32

  hm  10. oct. 2008 rev 1.3
    improved performance

  hm  18. oct. 2008 rev 1.4
    changed input en to e for compatibility reasons

  hm  10. mar. 2009 rev 1.5
    added type conversion for compatibility reasons
*)
END_FUNCTION_BLOCK

(* @PATH := '\/Mathematical\/functions' *)
FUNCTION_BLOCK FT_MIN_MAX
(*
  this function block stores the min and max value of an input signal.
  when rst is true the mn and mx outputs are set to the in value.
  when a rst is never active the function autoresets to the in value at startup.
  since the input might not be present at first cycle the mn and mx are set during second cycle.

  version 1.0 1 sep 2006
  programmer  hugo
  tested by   tobias
*)
  VAR_INPUT
    in : REAL;
    rst : BOOL;
  END_VAR
  VAR_OUTPUT
    mx : REAL;
    mn : REAL;
  END_VAR
  VAR
    init: BOOL;
  END_VAR

  IF rst OR NOT init THEN
    mn := in;
    mx := in;
    init := TRUE;
  ELSIF in < mn THEN mn := in;
  ELSIF in > mx THEN mx := in;
  END_IF;
END_FUNCTION_BLOCK

(* @PATH := '\/Mathematical\/functions' *)
FUNCTION_BLOCK FT_RMP
(*
  this ramp function follows an input signal with a linear ramp up or down, the up or down speed can be set with KF and KR.
  a K factor of 1 means 1 unit per second on the output. K factors can only be positive and not negative.
  a busy output signals the ramp is running or busy false means the in value is present on the output.
  a rmp input false means the output follows the input dierctly while a rmp = true means the output follows the input with a ramp.
  a updn output signal the directon of the ramp (up or down).

  version 1.4 25 jan 2008
  programmer  oscat
  tested by   oscat
*)
  VAR_INPUT
    Rmp : BOOL := TRUE;
    in : REAL;
    KR : REAL;
    KF : REAL;
  END_VAR
  VAR_OUTPUT
    out : REAL;
    busy : BOOL;
    UD : BOOL;
  END_VAR
  VAR
    tx: TIME;
    last: TIME;
    init: BOOL;
  END_VAR

  (* read system time *)
  tx := DWORD_TO_TIME(T_PLC_MS()) - last;

  IF NOT init THEN
    init := TRUE;
    last := tx;
    tx := t#0s;
    out := in;
  END_IF;
  IF NOT rmp THEN
    out := in;
    busy := FALSE;
  ELSIF out > in THEN
    (* ramp down *)
    out := out - TIME_TO_REAL(tx) * 0.001 * KF;
    out := MAX(in, out);
  ELSIF out < in THEN
    (* ramp up *)
    out := out + TIME_TO_REAL(tx) * 0.001 * KR;
    out := MIN(in, out);
  END_IF;

  (* set busy and dir flags *)
  IF out < in THEN
    busy := TRUE;
    ud := TRUE;
  ELSIF out > in THEN
    busy := TRUE;
    ud := FALSE;
  ELSE
    busy := FALSE;
  END_IF;
  last := last + tx;

(* revision history:
  hm 8.10.2006      rev 1.1
    added ud output

  hm 12. feb 2007   rev 1.2
    added init variable and corrected a possible startup problem

  hm  17. sep 2007  rev 1.3
    replaced time() with t_plc_ms() for compatibility reasons

  hm  25. jan 2008  rev 1.4
    performance improvements
    allow KR and KF to be 0
*)
END_FUNCTION_BLOCK

(* @PATH := '\/Mathematical\/functions' *)
FUNCTION LINEAR_INT : REAL
(*
  LINEAR_INT calculates an output based on a linear interpolation of up to 20 coordinates given in an array
  the input coordinates have to start at the lowest array position and must be sorted ba ascending X values.

  version 1.1 27 dec 2007
  programmer  oscat
  tested by   oscat
*)
  VAR_INPUT
    X : REAL;
    XY : OSCAT_BASIC_ARRAY1_20x0_1_OF_REAL; //ARRAY[1..20, 0..1] OF REAL;
    Pts : INT;
  END_VAR
  VAR
    i : INT;
  END_VAR

  (*make sure n is bound within the array size *)
  pts := MIN(pts,20);

  (* calculate the linear segement interpolation *)
  i := 2;
  (* search for segment and calculate output
    below and above the defined segments we interpolate the last segment *)
  WHILE (i < pts) AND (XY[i,0] < X) DO
    i := i + 1;
  END_WHILE;

  (* calculate the output value on the corresponding segment coordinates *)
  LINEAR_INT := ((XY[i,1] - XY[i-1,1]) * X - XY[i,1] * XY[i-1,0] + XY[i-1,1] * XY[i,0]) / (XY[i,0] - XY[i-1,0]);

(* revision history
  hm  7. oct 2007   rev 1.0
    original version

  hm  27 dec 2007   rev 1.1
    changed code for better performance
*)
END_FUNCTION

(* @PATH := '\/Mathematical\/functions' *)
FUNCTION POLYNOM_INT : REAL
(*
  POLYNOM_INT calculates an output based on a Polynom interpolation of up to 5 coordinates given in an array
  the indut coordinates have to start at the lowest array position and must be sorted ba ascending X values.

  version 1.3 10. mar. 2009
  programmer  oscat
  tested by   oscat
*)
  VAR_INPUT
    X : REAL;
    XY : ARRAY[1..5,0..1] OF REAL;
    Pts : INT;
  END_VAR
  VAR
    I, J : INT;
    stop: INT;
  END_VAR
  VAR_TEMP
    tmp : REAL;
  END_VAR

  (*make sure n is bound within the array size *)
  pts := MIN(pts, 5);

  (* this part is only to calculate the polynom parameters, which are then stores in the Y array
    the array values, it is not needed during runtime, unless the parameters will change during runtime
    the remaining code without this setup code can be used within a function to calculate specific functions
    the content of the arrays is then used as constant values within the function *)

  FOR i := 1 TO pts DO
    stop := i + 1;
      FOR j := pts TO stop BY -1 DO
        XY[j,1] := (XY[j,1] - XY[j-1,1]) / (XY[j,0] - XY[j-i,0]);
    END_FOR;
  END_FOR;

  (* this part is the actual calculation *)
  tmp := 0.0;
  FOR i := pts TO 1 BY -1 DO
         tmp := tmp * (X - XY[i,0]) + XY[i,1];
  END_FOR;
  POLYNOM_INT := tmp;

(* revision history
  hm  8. okt 2007 rev 1.0
    original version

  hm  17. dec 2007  rev 1.1
    init makes no sense for a function

  hm  22. feb 2008  rev 1.2
    improved performance

  hm  10. mar. 2009 rev 1.3
    changed syntax of real constants to 0.0
*)
END_FUNCTION

(* ---- Calculations.ST ---- *)
(* @PATH := '\/Engineering\/conversion' *)
FUNCTION_BLOCK ASTRO
(*
  this function converts different length units
  any unused input can simply be left open.
  different inputs connected at the same time will be added up.

  version 1.1 11. mar. 2009
  programmer  hugo
  tested by   oscat
*)
  VAR_INPUT
    m : REAL;
    AE : REAL;
    PC : REAL;
    LJ : REAL;
  END_VAR
  VAR_OUTPUT
    Ym : REAL;
    YAE : REAL;
    YPC : REAL;
    YLJ : REAL;
  END_VAR

  YAE :=  AE
      + m * 6.6845871535E-012
      + PC * 206265.0
      + LJ * 63240.0;
  Ym := YAE * 149.597870E9;
  YPC := YAE * 4.8481322570E-006;
  YLJ := YAE * 1.5812776724E-005;

(*
  Länge Meter m SI-Basiseinheit
  Astronomische Einheit* AE 1 AE = 149,597 870 · E9 m
  Parsec pc 1 pc = 206265 AE = 30,857 · E15 m
  Lichtjahr Lj 1 Lj = 9,460 530 · E15 m = 63240 AE = 0,306 59 pc
  Lngström L 1 L = E–l0 m
  typograph. Punkt p 1 p = 0,376 065 mm • im Druckereigewerbe
  inch** in 1 in = 2,54 · E–2 m = 25,4 mm***
  foot ft 1 ft = 0,3048 m = 30,48 cm
  yard yd 1 yd = 0,9144 m
  mile mile 1 mile = 1609,344 m
  Internat. Seemeile sm 1 sm = 1852 m
  Fathom fm 1 fm = 1,829 m • in der Seeschifffahrt
*)
(* revision history
  hm  27. mar. 2007 rev 1.0
    original version

  hm  11. mar. 2009 rev 1.1
    improved code
*)
END_FUNCTION_BLOCK

(* @PATH := '\/Engineering\/conversion' *)
FUNCTION BFT_TO_MS : REAL
(*
  this function converts wind speed from beaufort to m/s

  version 1.0 12. jun 2008
  programmer  hugo
  tested by   oscdat
*)
  VAR_INPUT
    BFT : INT;
  END_VAR

  BFT_TO_MS := EXPT( INT_TO_REAL(BFT), 1.5) * 0.836;

(* revision history
  hm  12. 6. 2008   rev 1.0
    original version
*)
END_FUNCTION

(* @PATH := '\/Engineering\/conversion' *)
FUNCTION C_TO_F : REAL
(*
  this function converts celsius  to fahrenheit

  version 1.1 11. mar. 2009
  programmer  hugo
  tested by   tobias
*)
  VAR_INPUT
    celsius : REAL;
  END_VAR

  C_TO_F := celsius * 1.8 + 32.0;

(* revision history
  hm  4. aug. 2006  rev 1.0
    original version

  hm  11. mar. 2009 rev 1.1
    real constants updated to new systax using dot
*)
END_FUNCTION

(* @PATH := '\/Engineering\/conversion' *)
FUNCTION C_TO_K : REAL
(*
  this function converts celsius to kelvin

  version 1.1 19. aug 2009
  programmer  hugo
  tested by   tobias
*)
  VAR_INPUT
    Celsius : REAL;
  END_VAR

  C_TO_K := Celsius - phys.T0;

(* revision history
  hm  4. aug 2006 rev 1.0
    original version

  hm  19. aug 2009  rev 1.1
    fixed calculation error
*)
END_FUNCTION

(* @PATH := '\/Engineering\/conversion' *)
FUNCTION DEG_TO_DIR : STRING[3]
(*
  this function converts degrees in compass direction.
  the function supports output in english (L=0) and german (L=1).

  version 1.1 22. oct. 2008
  programmer  hugo
  tested by   oscat
*)
  VAR_INPUT
    DEG : INT;
    N : INT;
    L : INT;
  END_VAR
  VAR
    ly: INT;
    word2 : WORD;
    word8 : WORD;
    tmp : INT;
  END_VAR

  IF L = 0 THEN ly := LANGUAGE.DEFAULT; ELSE ly := MIN(L, LANGUAGE.LMAX); END_IF;
  word2 := 2; word8 := 8;
  tmp := WORD_TO_INT(SHL(word2,INT_TO_UINT(N))) * WORD_TO_INT(SHR(word8,INT_TO_UINT(N)));
  DEG_TO_DIR := LANGUAGE.DIRS[ly, ((WORD_TO_INT(SHL(INT_TO_WORD(DEG),INT_TO_UINT(N-1))) + 45) / 90) MOD tmp];

(*
  DIR := ((SHL(DEG,N-1) + 45) / 90) MOD SHL(INT#2,N);
  explanation :
  DIR is calculated BY the following formula:
  DIR := ((DIR + 45) / 90) MOD 4 if N = 1 digit
  North = 0, East = 1 ....
  DIR := ((DIR + 22,5) / 45) MOD 8 if N = 2 digit
  convert to integer calculation
  DIR := ((DIR*2 + 45) / 90) MOD 8
  N = 0, NE = 1 ....
  ther above formula replaces 2^N with shift for performance
*)
(* revision histroy
  hm  11. jun. 2008 rev 1.0
    original release

  hm  22. oct. 2008 rev 1.1
    changed size of string variables to 30
*)
END_FUNCTION

(* @PATH := '\/Engineering\/conversion' *)
FUNCTION DIR_TO_DEG : INT
(*
  this function converts compass directions to degrees
  it will recognize up to 3 letter directions in english and german writing.

  version 1.1 22. oct. 2008
  programmer  hugo
  tested by oscat
*)
  VAR_INPUT
    DIR : STRING[3];
    L : INT;
  END_VAR
  VAR
    ly: INT;
    i : INT;
  END_VAR

  IF L = 0 THEN ly := LANGUAGE.DEFAULT; ELSE ly := MIN(L, LANGUAGE.LMAX); END_IF;
  FOR i := 0 TO 15 DO
    IF language.DIRS[ly, i] = DIR THEN EXIT; END_IF;
  END_FOR;
  DIR_TO_DEG := WORD_TO_INT(SHR(INT_TO_WORD(i * 45 + 1), 1));

(* revision histroy
  hm  22. oct. 2008 rev 1.1
    original release
*)
END_FUNCTION

(* @PATH := '\/Engineering\/conversion' *)
FUNCTION_BLOCK ENERGY
(*
  this function converts different energy units
  any unused input can simply be left open.
  different inputs connected at the same time will be added up.

  version 1.2 16. jan. 2010
  programmer  hugo
  tested by   oscat
*)
  VAR_INPUT
    J : REAL;
    C : REAL;
    Wh : REAL;
  END_VAR
  VAR_OUTPUT
    YJ : REAL;
    YC : REAL;
    YWh : REAL;
  END_VAR

  YJ := J + Wh * 3600.0 + C * 4.1868;
  YC := YJ * 0.238845896627496;
  YWh := YJ * 2.7777777778E-004;

(*
  Arbeit, Energie, Joule* J 1 J = 1 N · m = 1 W · s = (1/3,6) E–6 kW · h = 1 kg · m2/s2
  Wärmemenge Kilowattstunde kW · h 1 kW · h = 3,6 MJ = 860 kcal
  Elektronvolt eV 1 eV = 160,218 92 E–21 J
  Erg erg 1 erg = 1E–7 J
  Kalorie calorie 1 calalorie = 4,1868 J = 1,163 E–3 W · h
  Therm therm 1 therm = 105,50 · 106 J
*)
(* revision history
  hm  27. mar. 2007 rev 1.0
    original version

  hm  11. mar. 2009 rev 1.1
    improved code

  hm 16. jan 2010 rev 1.2
    avoid the string cal in comments for codesys import bug
*)
END_FUNCTION_BLOCK

(* @PATH := '\/Engineering\/conversion' *)
FUNCTION F_TO_C : REAL
(*
  this FUNCTION converts fahrenheit TO celsius

  version 1.1 11. mar. 2009
  programmer  hugo
  tested BY   tobias
*)
  VAR_INPUT
    fahrenheit : REAL;
  END_VAR

  F_TO_C := (fahrenheit - 32.0) * 0.5555555555555;

(* revision history
  hm  4. aug 2006 rev 1.0
    original version

  hm  11. mar. 2009 rev 1.1
    real constants updated to new systax using dot
*)
END_FUNCTION

(* @PATH := '\/Engineering\/conversion' *)
FUNCTION F_TO_OM : REAL
(*
  this function converts frequency to Omega F
  Omega = 2*PI*F

  version 1.1 18. oct. 2008
  programmer  hugo
  tested by oscat
*)
  VAR_INPUT
    F : REAL;
  END_VAR

  F_TO_OM := math.PI2 * F;

(* revision history
  hm  22. jan. 2007 rev 1.0
    original version

  hm  18. oct. 2008 rev 1.1
    unsing math constants
*)
END_FUNCTION

(* @PATH := '\/Engineering\/conversion' *)
FUNCTION F_TO_PT : TIME
(*
  this function converts frequency to periode time

  version 1.1 11. mar. 2009
  programmer  hugo
  tested by   tobias
*)
  VAR_INPUT
    F : REAL;
  END_VAR

  F_TO_PT := DWORD_TO_TIME(REAL_TO_DWORD(1.0 / F * 1000.0));

(* revision history
  hm  4. aug. 2006  rev 1.0
    original version

  hm  11. mar. 2009 rev 1.1
    real constants updated to new systax using dot
*)
END_FUNCTION

(* @PATH := '\/Engineering\/conversion' *)
FUNCTION GEO_TO_DEG : REAL
(*
  this function converts degrees, minutes seconds to decimal degrees.

  version 1.0 22. jan. 2009
  programmer  hugo
  tested by   oscat
*)
  VAR_INPUT
    D : INT;
    M : INT;
    SEC : REAL;
  END_VAR

  GEO_TO_DEG := INT_TO_REAL(D) + INT_TO_REAL(M) * 0.016666666666667 + sec * 0.00027777777777778;

(* revision histroy
   hm  22. jan. 2009 rev 1.0
   original release
*)
END_FUNCTION

(* @PATH := '\/Engineering\/conversion' *)
FUNCTION K_TO_C : REAL
(*
  this function converts kelvin to celsius

  version 1.1 19. aug 2009
  programmer  hugo
  tested by   tobias
*)
  VAR_INPUT
    Kelvin : REAL;
  END_VAR

  K_TO_C := Kelvin + phys.T0;

(* revision history
  hm  4. aug 2006 rev 1.0
    original version

  hm  19. aug 2009  rev 1.1
    fixed calculation error
*)
END_FUNCTION

(* @PATH := '\/Engineering\/conversion' *)
FUNCTION KMH_TO_MS : REAL
(*
  this function converts velocities from Kilometers / hour to Meters / Second

  version 1.1 6 jan 2007
  programmer  hugo
  tested by   tobias
*)
  VAR_INPUT
    kmh : REAL;
  END_VAR

  KMH_TO_MS := kmh * 0.2777777777777;

(* revision history
  hm  4. feb 2007   rev 1.0
    original version

  hm  6. jan 2008   rev 1.1
    improved performance
*)
END_FUNCTION

(* @PATH := '\/Engineering\/conversion' *)
FUNCTION_BLOCK LENGTH
(*
  this function converts different length units
  any unused input can simply be left open.
  different inputs connected at the same time will be added up.

  version 1.1 11. mar. 2009
  programmer  hugo
  tested by   oscat
*)
  VAR_INPUT
    m : REAL;
    p : REAL;
    in : REAL;
    ft : REAL;
    yd : REAL;
    mile : REAL;
    sm : REAL;
    fm : REAL;
  END_VAR
  VAR_OUTPUT
    Ym : REAL;
    Yp : REAL;
    Yin : REAL;
    Yft : REAL;
    Yyd : REAL;
    Ymile : REAL;
    Ysm : REAL;
    Yfm : REAL;
  END_VAR

  Ym := m
      + p * 0.000376065
      + in * 0.0254
      + ft * 0.3048
      + yd * 0.9144
      + mile * 1609.344
      + sm * 1852.0
      + fm * 1.829;
  Yp := Ym * 2659.11478068951;
  Yin := Ym * 39.37007874016;
  Yft := Ym * 3.28083989501;
  Yyd := Ym * 1.09361329834;
  Ymile := Ym * 0.00062137119;
  Ysm := Ym * 0.00053995680;
  Yfm := Ym * 0.54674685621;

(*
  Länge Meter m SI-Basiseinheit
  Astronomische Einheit* AE 1 AE = 149,597 870 · E9 m
  Parsec pc 1 pc = 206265 AE = 30,857 · E15 m
  Lichtjahr Lj 1 Lj = 9,460 530 · E15 m = 63240 AE = 0,306 59 pc
  Lngström L 1 L = E–l0 m
  typograph. Punkt p 1 p = 0,376 065 mm • im Druckereigewerbe
  inch** in 1 in = 2,54 · E–2 m = 25,4 mm***
  foot ft 1 ft = 0,3048 m = 30,48 cm
  yard yd 1 yd = 0,9144 m
  mile mile 1 mile = 1609,344 m
  Internat. Seemeile sm 1 sm = 1852 m
  Fathom fm 1 fm = 1,829 m • in der Seeschifffahrt
*)
(* revision history
  hm  27. mar. 2007 rev 1.0
    original version

  hm  11. mar. 2009 rev 1.1
    improved code
*)
END_FUNCTION_BLOCK

(* @PATH := '\/Engineering\/conversion' *)
FUNCTION MS_TO_BFT : INT
(*
  this function converts wind speed from M/s to beaufort

  version 1.0 12. jun 2008
  programmer  hugo
  tested by oscdat
*)
  VAR_INPUT
    MS : REAL;
  END_VAR

  MS_TO_BFT := REAL_TO_INT(EXPT(MS * 1.196172, 0.666667));

(* revision history
  hm  12. 6. 2008   rev 1.0
    original version
*)
END_FUNCTION

(* @PATH := '\/Engineering\/conversion' *)
FUNCTION MS_TO_KMH : REAL
(*
  this function converts velocities from Meters / Second to Kilometers / hour.

  version 1.0 4 Feb 2007
  programmer  hugo
  tested by   tobias
*)
  VAR_INPUT
    ms : REAL;
  END_VAR

  MS_TO_KMH := ms * 3.6;
END_FUNCTION

(* @PATH := '\/Engineering\/conversion' *)
FUNCTION OM_TO_F : REAL
(*
  this function converts Omega F to frequency
  F = OM / (2*PI)

  version 1.1 18. oct. 2008
  programmer  hugo
  tested by   tobias
*)
  VAR_INPUT
    OM : REAL;
  END_VAR

  OM_TO_F := OM / math.PI2;

(* revision history
  hm  22. jan. 2007 rev 1.0
    original version

  hm  18. oct. 2008 rev 1.1
    using math constants
*)
END_FUNCTION

(* @PATH := '\/Engineering\/conversion' *)
FUNCTION_BLOCK PRESSURE
(*
  this function converts different pressure units
  any unused input can simply be left open.
  different inputs connected at the same time will be added up.

  version 1.1 11. mar. 2009
  programmer  hugo
  tested by   oscat
*)
  VAR_INPUT
    mws : REAL;
    torr : REAL;
    att : REAL;
    atm : REAL;
    pa : REAL;
    bar : REAL;
  END_VAR
  VAR_OUTPUT
    Ymws : REAL;
    Ytorr : REAL;
    Yatt : REAL;
    Yatm : REAL;
    Ypa : REAL;
    Ybar : REAL;
  END_VAR

  Ybar := bar +
      pa * 1.0E-5 +
      0.980665 * att +
      1.01325 * atm +
      0.001333224 * torr +
      0.0980665 * mws;
  Ymws := ybar * 10.1971621297793;
  Ytorr := ybar * 750.0615050434140;
  Yatt := ybar * 1.0197162129779;
  yatm := ybar * 0.9869232667160;
  Ypa := ybar * 100000.0;

(*
  Druck, Pascal Pa 1 Pa = 1 N/m2 = 1 kg/(s2 �E m) . 0,75 �E 10.2 mmHg
  mechanische 1 MPa = 1 N/mm2 . fur Festigkeitsangaben
  Spannung Bar bar 1 bar = 105 Pa = 103 mbar = 105 kg/(s2 �E m)
  Millimeter- mmHg 1 mmHg = 133,322 Pa = 1,333 22 mbar
  Quecksilbersaule . nur in Heilkunde zulassig
  physik. Atmosphare atm 1 atm = 1,013 25 bar
  techn. Atmosphare at 1 at = 1 kp/cm2 = 0,980665 bar
  Torr Torr 1 Torr = (101325/760) Pa = 1,333224 mbar
  Meter-Wassersaule mWS 1 mWS = 9806,65 Pa = 98,0665 mbar
  psi lbf/in2 1 lbf/in2 = 68,947 57 mbar = 6894,757 Pa
*)
(* revision history
  hm  27. mar. 2007 rev 1.0
    original version

  hm  11. mar. 2009 rev 1.1
    improved code
*)
END_FUNCTION_BLOCK

(* @PATH := '\/Engineering\/conversion' *)
FUNCTION PT_TO_F : REAL
(*
  this function converts periode time to frequency

  version 1.1 11. mar. 2009
  programmer  hugo
  tested by   tobias
*)
  VAR_INPUT
    PT : TIME;
  END_VAR

  PT_TO_F := 1000.0 / DWORD_TO_REAL(TIME_TO_DWORD(PT));

(*  revision history
  hm  4. aug. 2006  rev 1.0
    original version

  hm  11. mar. 2009 rev 1.1
    real constants updated to new systax using dot
*)

END_FUNCTION

(* @PATH := '\/Engineering\/conversion' *)
FUNCTION_BLOCK SPEED
(*
  this function converts different speed units
  any unused input can simply be left open.
  different inputs connected at the same time will be added up.

  version 1.1 11. mar. 2009
  programmer  hugo
  tested by   oscat
*)
  VAR_INPUT
    ms : REAL;
    kmh : REAL;
    kn : REAL;
    mh : REAL;
  END_VAR
  VAR_OUTPUT
    Yms : REAL;
    Ykmh : REAL;
    Ykn : REAL;
    Ymh : REAL;
  END_VAR

  Yms := ms +
      kmh * 0.27777777777778 +
      kn * 0.5144444 +
      mh * 0.44704;
  Ykmh := Yms * 3.6;
  Ykn := Yms * 1.94384466037535;
  Ymh := Yms * 2.23693629205440;

(*
  Geschwindigkeit Meter durch Sekunde m/s 1 m/s = 3,6 km/h
  km durch (pro) Stunde, nicht „Stundenkilometer“ verwenden
  Knoten kn 1 kn = 1 sm/h = 0,5144 m/s
*)
(* revision history
  hm  27. mar. 2009 rev 1.0
    original version

  hm  11. mar. 2009 rev 1.1
    improved code
*)
END_FUNCTION_BLOCK

(* @PATH := '\/Engineering\/conversion' *)
FUNCTION_BLOCK TEMPERATURE
(*
  this function converts different temperature units
  any unused input can simply be left open.
  different inputs connected at the same time will be added up.

  version 1.0 21 feb 2008
  programmer  hugo
  tested by oscat
*)
  VAR_INPUT
    K : REAL;
    C : REAL := -273.15;
    F : REAL := -459.67;
    Re : REAL := -218.52;
    Ra : REAL;
  END_VAR
  VAR_OUTPUT
    YK : REAL;
    YC : REAL;
    YF : REAL;
    YRe : REAL;
    YRa : REAL;
  END_VAR

  YK := K + (C + 273.15) + (F + 459.67) * 0.555555555555 + (Re * 1.25 + 273.15) + (Ra * 0.555555555555);
  YC := YK -273.15;
  YF := YK * 1.8 - 459.67;
  YRe := (YK - 273.15) * 0.8;
  YRa := YK * 1.8;

(* revision history
  hm  21. feb. 2008 rev 1.0
    original version
*)
END_FUNCTION_BLOCK

(* ---- Control_Modules.ST ---- *)
(* @PATH := '\/Engineering\/control' *)
FUNCTION BAND_B : BYTE
(*
  BAND_B will limit X to B <= X <= 255-B. while X < B the resulkt will be 0 and while X > 255-B the output will be 255
  otherwise the result = X.

  version 1.0 21. Nov. 2008
  programmer  hugo
  tested by oscat
*)
  VAR_INPUT
    X : BYTE;
    B : BYTE;
  END_VAR

  IF X < B THEN
    BAND_B := 0;
  ELSIF BYTE_TO_USINT(X) > USINT#255 - BYTE_TO_USINT(B) THEN
    BAND_B := 255;
  ELSE
    BAND_B := X;
  END_IF;

(* revision history
  hm  21. nov. 2008 rev 1.0
    original version
*)
END_FUNCTION

(* @PATH := '\/Engineering\/control' *)
FUNCTION_BLOCK CONTROL_SET1
(*
  takahashi calculates controller parameters for P, PI and PID controllers based on the ziegler nichols method.

  version 1.1 11. mar. 2009
  programmer  hugo
  tested by   tobias
*)
  VAR_INPUT
    Kt : REAL;
    Tt : REAL;
    PI : BOOL;
    PID : BOOL;
  END_VAR
  VAR_INPUT //???CONSTANT
    P_K : REAL := 0.5;
    PI_K : REAL := 0.45;
    PI_TN : REAL := 0.83;
    PID_K : REAL := 0.6;
    PID_TN : REAL := 0.5;
    PID_TV : REAL := 0.125;
  END_VAR
  VAR_OUTPUT
    KP : REAL;
    TN : REAL;
    TV : REAL;
    KI : REAL;
    KD : REAL;
  END_VAR

  IF pi AND PID THEN
    KP := 0.0;
    TN := 0.0;
    TV := 0.0;
  ELSIF PID THEN
    KP := PID_K * Kt;
    TN := PID_TN * Tt;
    TV := PID_TV * Tt;
  ELSIF PI THEN
    KP := PI_K * Kt;
    TN := PI_TN * Tt;
  ELSE
    KP := P_K * Kt;
  END_IF;

  (* KI and KD are calculated *)
  IF tn > 0.0 THEN KI := KP / TN; ELSE KI := 0.0; END_IF;
  KD := KP * TV;

(* revision history
  hm  4. nov 2007 rev 1.0
    original version

  hm  11. mar. 2009 rev 1.1
  	real constants updated to new systax using dot
*)
END_FUNCTION_BLOCK

(* @PATH := '\/Engineering\/control' *)
FUNCTION_BLOCK CONTROL_SET2
(*
  takahashi calculates controller parameters for P, PI and PID controllers based on the ziegler nichols method.

  version 1.1 11. mar. 2009
  programmer  hugo
  tested by   tobias
*)
  VAR_INPUT
    KS : REAL;
    TU : REAL;
    TG : REAL;
    PI : BOOL;
    PID : BOOL;
  END_VAR
  VAR_INPUT //???CONSTANT
    P_K : REAL := 1.0;
    PI_K : REAL := 0.9;
    PI_TN : REAL := 3.33;
    PID_K : REAL := 1.2;
    PID_TN : REAL := 2.0;
    PID_TV : REAL := 0.5;
  END_VAR
  VAR_OUTPUT
    KP : REAL;
    TN : REAL;
    TV : REAL;
    KI : REAL;
    KD : REAL;
  END_VAR
  VAR
    TX : REAL;
  END_VAR

  IF TU > 0.0 AND KS > 0.0 THEN TX := TG / TU / KS; END_IF;
  IF pi AND PID THEN
    KP := 0.0;
    TN := 0.0;
    TV := 0.0;
  ELSIF PID THEN
    KP := PID_K * TX;
    TN := PID_TN * TU;
    TV := PID_TV * TU;
  ELSIF PI THEN
    KP := PI_K * TX;
    TN := PI_TN * TU;
  ELSE
    KP := P_K * TX;
  END_IF;

  (* KI and KD are calculated *)
  IF TN > 0.0 THEN KI := KP / TN; ELSE KI := 0.0; END_IF;
  KD := KP * TV;

(* revision history
  hm  4. nov 2007 rev 1.0
    original version

  hm  11. mar. 2009 rev 1.1
  	real constants updated to new systax using dot
*)
END_FUNCTION_BLOCK

(* @PATH := '\/Engineering\/control' *)
FUNCTION DEAD_ZONE : REAL
(*
  dead_zone2 is a linear transfer function which follows a linear function except for x is close to 0.
  Y = X if abs(x) > L otherwise its 0.

  version 1.2 11. mar. 2009
  programmer  hugo
  tested by   oscat
*)
  VAR_INPUT
    X : REAL;
    L : REAL;
  END_VAR

  IF ABS(x) > L THEN
    dead_zone := X;
  ELSE
    DEAD_ZONE := 0.0;
  END_IF;

(* revision history
  hm  12. feb. 2007 rev 1.0
    original version

  hm  14. jun. 2008 rev 1.1
    improved performance

  hm  11. mar. 2009 rev 1.2
    real constants updated to new systax using dot
*)
END_FUNCTION

(* @PATH := '\/Engineering\/control' *)
FUNCTION CTRL_IN : REAL
(*

  version 1.0 2. jun 2008
  programmer  hugo
  tested by   tobias
*)
  VAR_INPUT
    SET_POINT, ACTUAL, NOISE : REAL;
  END_VAR

  (* calculate the process error DIFF *)
  CTRL_IN := DEAD_ZONE(SET_POINT - ACTUAL, NOISE);

(* revision history
  hm  2. jun. 2008  rev 1.0
    original version
*)
END_FUNCTION

(* @PATH := '\/Engineering\/control' *)
FUNCTION_BLOCK CTRL_OUT
(*

  version 1.1 5. nov 2008
  programmer  hugo
  tested by oscat
*)
  VAR_INPUT
    CI, OFFSET, MAN_IN, LIM_L, LIM_H : REAL;
    MANUAL : BOOL;
  END_VAR
  VAR_OUTPUT
    Y : REAL;
    LIM : BOOL;
  END_VAR

  Y := SEL(MANUAL, CI, MAN_IN) + OFFSET;

  (* Limit the output *)
  IF Y > LIM_L AND Y < LIM_H THEN
    LIM := FALSE;
  ELSE
    Y := LIMIT(LIM_L, Y, LIM_H);
    LIM := TRUE;
  END_IF;

(* revision history
  hm  2. jun. 2008  rev 1.0
    original version

  hm  5. nov. 2008  rev 1.1
    optimized code
*)
END_FUNCTION_BLOCK

(* @PATH := '\/Engineering\/control' *)
FUNCTION_BLOCK FT_PIWL
(*
  FT_PIWL is a PI controller.
  The PID controller works according to the fomula Y = IN *(KP+ KI * INTEG(e) ).
  a rst will reset the integrator to 0
  lim_h and Lim_l set the possible output range of the controller.
  the output flag lim will signal that the output limits are active.
  the integrator ist equipped with anti wind-up circuitry which limits trhe total output ranke to lim_l and lim_h

  default values for KP = 1, KI = 1, ILIM_L = -1E37, iLIM_H = +1E38.
  version 1.3 11. mar. 2009
  programmer  hugo
  tested by   oscat
*)
  VAR_INPUT
    IN : REAL;
    KP : REAL := 1.0;
    KI : REAL := 1.0;
    LIM_L : REAL := -1.0E38;
    LIM_H : REAL := 1.0E38;
    RST : BOOL;
  END_VAR
  VAR_OUTPUT
    Y : REAL;
    LIM : BOOL;
  END_VAR
  VAR
    init: BOOL;
    tx: UDINT; //DWORD;
    tc : REAL;
    t_last: UDINT; //DWORD;
    in_last : REAL;
    i: REAL;
    p: REAL;
  END_VAR

  (* initialize at power_up *)
  IF NOT init OR RST THEN
    init := TRUE;
    in_last := in;
    t_last := DWORD_TO_UDINT( T_PLC_US());
    i := 0.0;
    tc := 0.0;
  ELSE
    (* read last cycle time in Microseconds *)
    tx := DWORD_TO_UDINT( T_PLC_US());
    tc := UDINT_TO_REAL(tx - t_last);
    t_last := tx;

    (* calculate proportional part *)
    p := KP * IN;

    (* run integrator *)
    i := (IN + in_last) * 5.0E-7 * KI * tc + i;
    in_last := IN;

    (* calculate output Y *)
    Y := p + i;

    (* check output for limits *)
    IF Y >= LIM_H THEN
      Y := LIM_H;
      IF ki <> 0.0 THEN
        i := LIM_H - p;
      ELSE
        i := 0.0;
      END_IF;
      LIM := TRUE;
    ELSIF Y <= LIM_L THEN
      Y := LIM_L;
      IF ki <> 0.0 THEN
        i := LIM_L - p;
      ELSE
        i := 0.0;
      END_IF;
      LIM := TRUE;
    ELSE
      LIM := FALSE;
    END_IF;
  END_IF;

(* revision history
  hm 13. jun. 2008  rev 1.0
    original version

  hm  27. oct. 2008 rev 1.1
    integrator will not be adjusted when ki = 0

  hm  25. jan 2009  rev 1.2
    module will also work with negative K

  hm  11. mar. 2009 rev 1.3
    real constants updated to new systax using dot
*)
END_FUNCTION_BLOCK

(* @PATH := '\/Engineering\/control' *)
FUNCTION_BLOCK CTRL_PI
(*
  FT_PI is a PI controller with manual functionality.
  The PID controller works according to the fomula Y = e *(KP+ KI * INTEG(e) ) + offset, while e = set_point - actual.
  a rst will reset all internal data, while a switch to manual will cause the controller to follow the function Y = manual_in + offset.
  limit_h and Limit_l set the possible output range of Y.
  the output flags lim will signal that the output limits are active and overflow will signal that the integrator has reached its limits.

  since rev 1.1 the "trapezregel is used for more accuracy.
  rev 1.2 added selective integratin which means the integrative component is only active within a small range of the target value
  this avoids the integrator to go to limits while an input setpoint change happened and is only causing overshoots.
  the int_band is by default 100 which means the int is active all the time and if set to for example to 0.1 the integrator is only active
  while the input is between 0.9 and 1.1 of the set_point value.

  default values for KP = 1, TN = 1, TV = 1, LIMIT_L = -1000, LIMIT_H = +1000.
  version 2.0 30. jun 2008
  programmer  hugo
  tested by oscat
*)
  VAR_INPUT
    ACT, SET, SUP, OFS, M_I : REAL;
    MAN : BOOL;
    RST : BOOL;
    KP : REAL := 1.0;
    KI : REAL := 1.0;
    LL : REAL := -1000.0;
    LH : REAL := 1000.0;
  END_VAR
  VAR_OUTPUT
    Y : REAL;
    DIFF : REAL;
    LIM : BOOL;
  END_VAR
  VAR
    pi : FT_PIWL;
    co : CTRL_OUT;
  END_VAR

  DIFF := CTRL_IN(SET, ACT, SUP);
  pi(in := DIFF, kp := KP, ki := KI, lim_l := LL, lim_h := LH, rst := RST);
  co(ci := pi.Y, OFFSET := OFS, man_in := M_I, lim_l := LL, lim_h := LH, MANUAL := MAN);
  Y := co.Y;
  LIM := co.LIM;

(* revision history
  hm  31.10.2007    rev 1.0
    original version

  hm  3.11.2007   rev 1.1
    added noise input to filter noise
    added output diff
    set limit output false when output is within limits
    overfolw was not set correctly

  hm  5. jan 2008   rev 1.2
    improved performance

  hm  20. jun. 2008 rev 2.0
    rewritten using new modular approach
*)
END_FUNCTION_BLOCK

(* @PATH := '\/Engineering\/control' *)
FUNCTION_BLOCK FT_DERIV
(*
  FT_deriv calculates the derivate over the signal "in" with Faktor "K".
  a run input enables or stops the calculation, if left unconnected its true and therfore the calculation is executed.
  if K is not specified the default is 1.

  version 1.5 11. mar. 2009
  programmer  hugo
  tested by   oscat
*)
  VAR_INPUT
    in : REAL;
    K : REAL := 1.0;
    run : BOOL := TRUE;
  END_VAR
  VAR_OUTPUT
    out : REAL;
  END_VAR
  VAR
    old: REAL;
    tx: UDINT; //DWORD;
    last: UDINT; //DWORD;
    init: BOOL;
    tc: REAL;
  END_VAR

  (* read system time *)
  tx := DWORD_TO_UDINT(T_PLC_US());
  tc := UDINT_TO_REAL(tx - last);
  last := tx;

  (* init on first startup *)
  IF NOT init THEN
    init := TRUE;
    old := in;
  ELSIF run AND tc > 0.0 THEN
    out := (in - old) / tc * 1000000.0 * K;
    old := in;
  ELSE
    out := 0.0;
  END_IF;

(*
  hm 3.1.2007     rev 1.1
    added init code for startup
    set the default for K to 1

  hm  15. sep 2007  rev 1.2
    replaced Time() with T_PLC_US for compatibility and performance reasons
    increased accuracy and work in microseconds internally

  hm 29 oct 2007  rev 1.3
    prohibit calculation when tx - last = 0 to avoid division by 0 and increase accuracy on fast systems

  hm  6. nov. 2008  rev 1.4
    improved performance

  hm  11. mar. 2009 rev 1.5
    inproved code
*)
END_FUNCTION_BLOCK

(* @PATH := '\/Engineering\/control' *)
FUNCTION_BLOCK FT_PIDWL
(*
  FT_PIDWL is a PID controller with dynamic wind_up reset.
  The PID controller works according to the fomula Y = KP *(IN + KI * INTEG(e) + DERIV(e) ).
  a rst will reset the integrator to 0
  lim_h and Lim_l set the possible output range of the internal integrator.
  the output flags lim will signal that the output limits are active.

  default values for KP = 1, KI = 1, ILIM_L = -1E37, iLIM_H = +1E38.
  version 1.3 13. nov. 2009
  programmer  hugo
  tested by   tobias
*)
  VAR_INPUT
    IN : REAL;
    KP : REAL := 1.0;
    TN : REAL := 1.0;
    TV : REAL := 1.0;
    LIM_L : REAL := -1.0E38;
    LIM_H : REAL := 1.0E38;
    RST : BOOL;
  END_VAR
  VAR_OUTPUT
    Y : REAL;
    LIM : BOOL;
  END_VAR
  VAR
    piwl : FT_PIWL;
    diff : FT_DERIV;
  END_VAR

  (* if rst then *)
  IF rst THEN
    piwl(rst := TRUE);
    piwl.RST := FALSE;
  ELSE
    (* run PIWL controller first *)
    (* we need to check if TN = 0 and do alternative calls *)
    IF TN = 0.0 THEN
      piwl(in := IN * KP, KP := 1.0, KI := 0.0, LIM_L := LIM_L, LIM_H := LIM_H);
    ELSE
      piwl(in := IN * KP, KP := 1.0, KI := 1.0 / TN, LIM_L := LIM_L, LIM_H := LIM_H);
    END_IF;

    (* run differentiator and add_to_output *)
    diff(IN := IN, K := KP * TV);
    Y := piwl.Y + diff.out;

    (* limit the output *)
    IF Y < LIM_L THEN
      LIM := TRUE;
      Y := LIM_L;
    ELSIF Y > LIM_H THEN
      LIM := TRUE;
      Y := LIM_H;
    ELSE
      LIM := FALSE;
    END_IF;
  END_IF;

(* revision history
  hm 13. jun. 2008  rev 1.0
    original version

  hm  25. jan 2008  rev 1.1
    multiply differential part with KP

  hm  11. mar. 2009 rev 1.2
    real constants updated to new systax using dot

  hm  13. nov. 2009 rev 1.3
    fixed code for negative KP
*)
END_FUNCTION_BLOCK

(* @PATH := '\/Engineering\/control' *)
FUNCTION_BLOCK CTRL_PID
(*
  FT_PI is a PI controller with manual functionality.
  The PID controller works according to the fomula Y = e *(KP+ KI * INTEG(e) ) + offset, while e = set_point - actual.
  a rst will reset all internal data, while a switch to manual will cause the controller to follow the function Y = manual_in + offset.
  limit_h and Limit_l set the possible output range of Y.
  the output flags lim will signal that the output limits are active.

  version 2.0 30. jun. 2008
  programmer  hugo
  tested by oscat
*)
  VAR_INPUT
    ACT, SET, SUP, OFS, M_I : REAL;
    MAN : BOOL;
    RST : BOOL;
    KP : REAL := 1.0;
    TN : REAL := 1.0;
    TV : REAL := 1.0;
    LL : REAL := -1000.0;
    LH : REAL := 1000.0;
  END_VAR
  VAR_OUTPUT
    Y : REAL;
    DIFF : REAL;
    LIM : BOOL;
  END_VAR
  VAR
    pid : FT_PIDWL;
    co : CTRL_OUT;
  END_VAR

  DIFF := CTRL_IN(SET, ACT, SUP);
  pid(in := DIFF, kp := KP, tn := TN, tv := TV, lim_l := LL, lim_h := LH, rst := RST);
  co(ci := pid.Y, OFFSET := OFS, man_in := M_I, lim_l := LL, lim_h := LH, MANUAL := MAN);
  Y := co.Y;
  LIM := co.LIM;

(* revision history
  hm 1.12.2006    rev 1.1
    changed algorithm to trapezregel for higher accuracy.

  hm 3.1.2007   rev 1.2
    added integ_band to select when the integrator is active.

  hm  3.3.2007    rev 1.3
    added default values to inputs KP, TN, TV, LIMIT_L und LIMIT_H.

  hm 31.oct 2007  rev 1.4
    total rewrite of the module to avoid failures when one of the limits is 0

  hm  3.11.2007 rev 1.5
    added noise input to filter noise
    added output diff
    set limit output false when output is within limits
    overfolw was not set correctly

  hm  5. jan 2008 rev 1.6
    improved code for better performance
*)
END_FUNCTION_BLOCK

(* @PATH := '\/Engineering\/control' *)
FUNCTION_BLOCK CTRL_PWM
(*

  version 1.1 21. oct. 2008
  programmer  hugo
  tested by oscat
*)
  VAR_INPUT
    CI, MAN_IN : REAL;
    MANUAL : BOOL;
    F : REAL;
  END_VAR
  VAR_OUTPUT
    Q : BOOL;
  END_VAR
  VAR
    PW : PWM_DC;
  END_VAR

  PW(F := F, DC := SEL(MANUAL,CI,MAN_IN));
  Q := PW.Q;

(* revision history
  hm 3. jun. 2008   rev 1.0
    original version

  hm  21. oct. 2008 rev 1.1
    optimized code
*)
END_FUNCTION_BLOCK

(* @PATH := '\/Engineering\/control' *)
FUNCTION DEAD_BAND : REAL
(*
  DEAD_BAND ist eine lineare Übertragungsfunktion mit Totzone. Die Funktion verschiebt den positiven Teil der Kurve um +L und den negativen Teil der Kurve um -L.
  DEAD_BAND = X - L wenn X > L)
  DEAD_BAND = X + L wenn X < -L
  DEAD_BAND = 0 wenn Abs(X) <= L

  version 1.2 18. jan. 2011
  programmer  hugo
  tested by   oscat
*)
  VAR_INPUT
    X : REAL;
    L : REAL;
  END_VAR

  IF X > L THEN
    DEAD_BAND := X - L;
  ELSIF X < -L THEN
    DEAD_BAND := X + L;
  ELSE
    DEAD_BAND := 0.0;
  END_IF;

(* revision history
  hm  2. nov. 2007  rev 1.0
    original version

  hm  14. jun. 2008 rev 1.1
    improved performance

  hm  18. jan. 2011 rev 1.2
    assign 0 before return
*)
END_FUNCTION

(* @PATH := '\/Engineering\/control' *)
FUNCTION_BLOCK FT_PT1
(*
  FT_PT1 is an low pass filter with a programmable time T and faktor K.

  version 1.11  18. jan. 2011
  programmer  hugo
  tested by   oscat
*)
  VAR_INPUT
    in : REAL;
    T : TIME;
    K : REAL := 1.0;
  END_VAR
  VAR_OUTPUT
    out : REAL;
  END_VAR
  VAR
    last : UDINT; //DWORD;
    tx: UDINT; //DWORD;
    init: BOOL;
  END_VAR

  (* read system time *)
  tx := DWORD_TO_UDINT( T_PLC_US());

  (* startup initialisation *)
  IF NOT init OR T = t#0s THEN
    init := TRUE;
    out := K * in;
  ELSE
    out := out + (in * K - out) * UDINT_TO_REAL(Tx - last) / TIME_TO_REAL(T) * 1.0E-3;
    IF ABS(out) < 1.0E-20 THEN out := 0.0; END_IF;
  END_IF;
  last := tx;

(*
  hm 1.1.2007 rev 1.1
    corrected error while startup value was not correct
    for very small time values real output would run out of range.

  hm 3.1.2007 rev 1.2
    corrected an error for falling edge failures.
    added output faktor K.

  hm 27. 2. 2007  rev 1.3
    output will be input during init for definitive startup condition.

  hm  15.9.2007 rev 1.4
    changed time() to T_PLC_US() for compatibilitxy resons
    increased internal accuracy to Microseconds instead of Milliseconds

  hm  23. oct 2007  rev 1.5
    added out := in to the init statements

  hm  30. nov 2007  rev 1.6
    changed out to be K * in during initialization

  hm  5. jan 2008 rev 1.7
    improved code for better performance

  hm  16. mar. 2008 rev 1.8
    added type conversion to avoid warning under codesys 3.0

  hm  14. jun. 2008 rev 1.9
    improved code

  hm  11. mar. 2009 rev 1.10
    real constants updated to new systax using dot

  hm  18. jan. 2011 rev 1.11
    avoid underrun of out
*)
END_FUNCTION_BLOCK

(* @PATH := '\/Engineering\/control' *)
FUNCTION_BLOCK DEAD_BAND_A
(*
  DEAD_BAND ist eine lineare Übertragungsfunktion mit Totzone. Die Funktion verschiebt den positiven Teil der Kurve um -L und den negativen Teil der Kurve um +L.
  DEAD_BAND = X wenn Abs(X) > L wenn Abs(X) > L
  DEAD_BAND = 0 wenn Abs(X) <= L
  Die Breite der Totzone wird automatisch aus dem Signalrauschen errechnet.

  version 1.1 11. mar. 2009
  programmer  hugo
  tested by   oscat
*)
  VAR_INPUT
    X : REAL;
    T : TIME;
    KL : REAL := 1.0;
    LM : REAL;
  END_VAR
  VAR_OUTPUT
    Y : REAL;
    L : REAL;
  END_VAR
  VAR
    tp1 : FT_PT1;
    tp2 : FT_PT1;
  END_VAR

  (* filter the input signal *)
  tp1(in := X, T:= T);

  (* filter the HF portion to generate a stable L *)
  tp2(in := ABS(tp1.out - X), T := MULTIME(T, 4.0));

  (* now we determine L which is half the width of the dead band *)
  L := MIN(KL * tp2.out, LM);

  IF X > L THEN
    Y := X - L;
  ELSIF X < -L THEN
    Y := X + L;
  ELSE
    Y := 0.0;
  END_IF;

(* revision history
  hm  14. jun. 2008 rev 1.0
    original version

  hm  11. mar. 2009 rev 1.1
    real constants updated to new systax using dot
*)
END_FUNCTION_BLOCK

(* @PATH := '\/Engineering\/control' *)
FUNCTION_BLOCK DEAD_ZONE2
(*
  dead_zone2 is a linear transfer function which follows a linear function except for x is close to 0.
  Y = X if abs(x) > L.
  for values of 0 +/- L a hysteresis function will hold the output at + or - L.

  version 1.1 11. mar. 2009
  programmer  hugo
  tested by   tobias
*)
  VAR_INPUT
    X : REAL;
    L : REAL;
  END_VAR
  VAR_OUTPUT
    Y: REAL;
  END_VAR

  IF ABS(x) > L THEN
    Y := X;
  ELSIF Y > 0.0 THEN
    Y := L;
  ELSE
    Y := -L;
  END_IF;

(* revision history
  hm  12. feb. 2007 rev 1.0
    original version

  hm  11. mar. 2009 rev 1.1
    real constants updated to new systax using dot
*)
END_FUNCTION_BLOCK

(* @PATH := '\/Engineering\/control' *)
FUNCTION_BLOCK FT_IMP
(*
  FT_IMP is   an impulse filter (high pass filter) with the time T and factor K.

  version 1.1 3 Jan 2007
  programmer  hugo
  tested by oscat
*)
  VAR_INPUT
    in : REAL;
    T : TIME;
    K : REAL := 1.0;
  END_VAR
  VAR_OUTPUT
    out : REAL;
  END_VAR
  VAR
    t1 : FT_PT1;
  END_VAR

  T1(in:= in, T:=T);
  out := (in - t1.out) * K;

(*
  hm 3.1.2007 rev 1.1
    added factor K
*)
END_FUNCTION_BLOCK

(* @PATH := '\/Engineering\/control' *)
FUNCTION_BLOCK INTEGRATE
(*
  integrate is a plain integrator with I/O for out.

  version 1.0 3. nov. 2008
  programmer  hugo
  tested by oscat
*)
  VAR_INPUT
    E : BOOL := TRUE;
    X : REAL;
    K : REAL := 1.0;
  END_VAR
  VAR_IN_OUT
    Y : REAL;
  END_VAR
  VAR
    X_last : REAL;
    init: BOOL;
    last: UDINT; //DWORD;
    tx: UDINT; //DWORD;
  END_VAR

  (*read system time *)
  tx := DWORD_TO_UDINT( T_PLC_MS());

  IF NOT init THEN
    init := TRUE;
    X_last := X;
  ELSIF E THEN
    Y := (X + X_LAST) * 0.5E-3 * UDINT_TO_REAL(tx-last) * K + Y;
    X_last := X;
  END_IF;
  last := tx;

(*
  hm 3. nov. 2008 rev 1.0
  original version
*)
END_FUNCTION_BLOCK

(* @PATH := '\/Engineering\/control' *)
FUNCTION_BLOCK FT_INT
(*
  FT_int is an integrator with input IN and factor K.
  integration is only done while run = true, if run is false integration is stopped and the out remains at the last value.
  if run is left unconnected, run is considered true by the function block.
  the output ET will display the total integration time from last reset.
  the out_min and out_max values can be set to ,imit the output value range.
  the default for K is 1.

  version 2.2 10. mar. 2009
  programmer  hugo
  tested by   oscat
*)
  VAR_INPUT
    IN : REAL;
    K : REAL := 1;
    RUN : BOOL := TRUE;
    RST : BOOL;
    OUT_MIN : REAL := -1E37;
    OUT_MAX : REAL := 1E37;
  END_VAR
  VAR_OUTPUT
    OUT : REAL;
    LIM : BOOL;
  END_VAR
  VAR
    INTeg : INTEGRATE;
  END_VAR

  IF rst THEN
    out := 0.0;
  ELSE
    integ(X := IN, E := RUN, K := K, Y := out);
  END_IF;

  (* limit the outputs *)
  IF out >= OUT_MAX THEN
    out := out_max;
    LIM := TRUE;
  ELSIF out <= out_min THEN
    out := out_min;
    lim := TRUE;
  ELSE
    lim := FALSE;
  END_IF;

(*
  hm 13.12.2006 rev 1.1
    changed to "trapezregel" which increases accuracy
    before out := out + in * time new: out := out + (in + in_last) / 2 * time

  hm 15.1.2007    rev 1.2
    added default for k to be 1.

  hm  15.9.2007   rev 1.3
    replaced time() with T_PLC_US for compatibility and performance reason
    increased internal accuracy to microseconds

  hm 29. oct 2007   rev 1.4
    changed code so int will not be called is time difference is 0 to increase accuracy on systems
    with cycle times below 1ms

  hm  2. dec 2007   rev 1.5
    changed code for better performance

  hm  5. jan 2008   rev 1.6
    further improvements in performance

  hm  8. feb 2008   rev 1.7
    deleted limits +/- 1000 now limit is the range of real
    added variables out1 and out2 to extend the resolution
    corrected an error with elapsed time
    deleted unusfull output ET

  hm  13. mar 2008  rev 1.8
    changed preset value out_min to -1e37.
    stop integrator at the limits.

  hm  16. mar 2008  rev 1.9
    added type conversion to avoid warning under codesys 3.0

  hm  2. jun. 2008  rev 2.0
    rewritten with clear code
    limits can now be set without run

  hm  3. nov. 2008  rev 2.1
    optimized code using INTEGRATE and LIMX

  hm  10. mar. 2009 rev 2.2
    removed nested comments
*)
END_FUNCTION_BLOCK

(* @PATH := '\/Engineering\/control' *)
FUNCTION_BLOCK FT_INT2
(*
  FT_int2 is an integrator with input IN and factor K.
  integration is only done while run = true, if run is false integration is stopped and the out remains at the last value.
  if run is left unconnected, run is considered true by the function block.
  the out_min and out_max values can be set to ,imit the output value range.
  the default for K is 1.
  FT_INT2 has double presision accuracy (14 digits).

  version 1.2 11. mar. 2009
  programmer  hugo
  tested by   oscat
*)
  VAR_INPUT
    IN : REAL;
    K : REAL := 1.0;
    RUN : BOOL := TRUE;
    RST : BOOL;
    OUT_MIN : REAL := -1.0E38;
    OUT_MAX : REAL := 1.0E38;
  END_VAR
  VAR_OUTPUT
    OUT : REAL;
    LIM : BOOL;
  END_VAR
  VAR
    integ: INTEGRATE;
    ix : REAL;
    val : REAL2;
  END_VAR

  IF RST THEN
    val := R2_SET(0.0);
    out := 0.0;
  ELSE
    integ(X := IN, E := RUN, K := K, Y := ix);
    val := R2_ADD(val, ix);
    ix := 0.0;
    OUT := val.RX;
  END_IF;

  (* check output for limits *)
  IF out > OUT_MIN AND out < OUT_MAX THEN
    LIM := FALSE;
  ELSE
    OUT := LIMIT(OUT_MIN, OUT, OUT_MAX);
    val := R2_SET(OUT);
    LIM := TRUE;
  END_IF;

(*  revision history
  hm  2. jun. 2008  rev 1.0
    original version

  hm  5. nov. 2008  rev 1.1
    rewritten code using integrate

  hm  11. mar. 2009 rev 1.2
    real constants updated to new systax using dot
*)
END_FUNCTION_BLOCK

(* @PATH := '\/Engineering\/control' *)
FUNCTION_BLOCK FT_PD
(*
  FT_PD is a PD controller.
  The PD controller works according to the fomula Y = KP *(IN + DERIV(e) ).

  version 1.0 3. jun 2008
  programmer  hugo
  tested by   tobias
*)
  VAR_INPUT
    IN : REAL;
    KP : REAL := 1.0;
    TV : REAL := 1.0;
  END_VAR
  VAR_OUTPUT
    Y : REAL;
  END_VAR
  VAR
    diff : FT_DERIV;
  END_VAR

  (* run differentiator *)
  diff(IN := IN, K := TV);

  (* combine both values *)
  Y := KP * (diff.out + IN);

(* revision history
  hm  3. jun. 2008  rev 1.0
    original version
*)
END_FUNCTION_BLOCK

(* @PATH := '\/Engineering\/control' *)
FUNCTION_BLOCK FT_PDT1
(*
  FT_PD is a PD controller.
  The PD controller works according to the fomula Y = KP *(IN + DERIV(e) ).

  version 1.0 3. jun 2008
  programmer  hugo
  tested by   tobias
*)
  VAR_INPUT
    IN : REAL;
    KP : REAL := 1.0;
    TV : REAL := 1.0;
    T1 : REAL := 1.0;
  END_VAR
  VAR_OUTPUT
    Y : REAL;
  END_VAR
  VAR
    diff : FT_DERIV;
    TP : FT_PT1;
  END_VAR

  (* run differentiator *)
  diff(IN := IN, K := TV);

  (* Run PT1 filter *)
  tp(in := diff.out, T := REAL_TO_TIME(T1));

  (* combine both values *)
  Y := KP * (tp.out + IN);

(* revision history
  hm  3. jun. 2008  rev 1.0
    original version
*)
END_FUNCTION_BLOCK

(* @PATH := '\/Engineering\/control' *)
FUNCTION_BLOCK FT_PI
(*
  FT_PI is a PI controller.
  The PID controller works according to the fomula Y = IN *(KP+ KI * INTEG(e) ).
  a rst will reset the integrator to 0
  ilim_h and iLim_l set the possible output range of the internal integrator.
  the output flags lim will signal that the output limits are active.

  default values for KP = 1, KI = 1, ILIM_L = -1E37, iLIM_H = +1E38.
  version 2.0 3. jun 2008
  programmer  hugo
  tested by   tobias
*)
  VAR_INPUT
    IN : REAL;
    KP : REAL := 1.0;
    KI : REAL := 1.0;
    ILIM_L : REAL := -1E38;
    ILIM_H : REAL := 1E38;
    IEN : BOOL := TRUE;
    RST : BOOL;
  END_VAR
  VAR_OUTPUT
    Y : REAL;
    LIM : BOOL;
  END_VAR
  VAR
    integ : FT_INT;
  END_VAR

  (* run integrator *)
  integ(IN := IN, K := KI, RUN := IEN, RST := RST, OUT_MIN := ILIM_L, OUT_MAX := ILIM_H);

  (* check if integrator has reached its limits and set overflow *)
  LIM := integ.LIM;
  Y := KP * IN + integ.Out;

(* revision history
  hm  3. jun. 2008  rev 2.0
    original version
*)
END_FUNCTION_BLOCK

(* @PATH := '\/Engineering\/control' *)
FUNCTION_BLOCK FT_PID
(*
  FT_PI is a PI controller.
  The PID controller works according to the fomula Y = IN *(KP+ KI * INTEG(e) ).
  a rst will reset the integrator to 0
  ilim_h and iLim_l set the possible output range of the internal integrator.
  the output flags lim will signal that the output limits are active.

  default values for KP = 1, KI = 1, ILIM_L = -1E37, iLIM_H = +1E38.
  version 2.1 11. mar. 2009
  programmer  hugo
  tested by   tobias
*)
  VAR_INPUT
    IN : REAL;
    KP : REAL := 1.0;
    TN : REAL := 1.0;
    TV : REAL := 1.0;
    ILIM_L : REAL := -1.0E38;
    ILIM_H : REAL := 1.0E38;
    IEN : BOOL := TRUE;
    RST : BOOL;
  END_VAR
  VAR_OUTPUT
    Y : REAL;
    LIM : BOOL;
  END_VAR
  VAR
    integ : FT_INT;
    diff : FT_DERIV;
  END_VAR

  (* run integrator only if TN > 0 *)
  IF TN > 0.0 THEN
    integ(IN := IN, K := 1.0 / TN, RUN := IEN, RST := RST, OUT_MIN := ILIM_L, OUT_MAX := ILIM_H);
  ELSE
    integ(RST := FALSE);
  END_IF;

  (* run differentiator *)
  diff(IN := IN, K := TV);

  (* combine both values *)
  Y := KP * (integ.Out + diff.out + IN);

  (* check if integrator has reached its limits and set overflow *)
  LIM := integ.LIM;

(* revision history
  hm 3. jun. 2008   rev 2.0
    original version

  hm  11. mar. 2009 rev 2.1
    real constants updated to new systax using dot
*)
END_FUNCTION_BLOCK

(* @PATH := '\/Engineering\/control' *)
FUNCTION_BLOCK FT_PIDW
(*
  FT_PIDW is a PID controller with dynamic wind_up reset.
  The PID controller works according to the fomula Y = KP *(IN + KI * INTEG(e) + DERIV(e) ).
  a rst will reset the integrator to 0
  lim_h and Lim_l set the possible output range of the internal integrator.
  the output flags lim will signal that the output limits are active.

  default values for KP = 1, KI = 1, ILIM_L = -1E37, iLIM_H = +1E38.
  version 1.2 11. mar. 2009
  programmer  hugo
  tested by   oscat
*)
  VAR_INPUT
    IN : REAL;
    KP : REAL := 1.0;
    TN : REAL := 1.0;
    TV : REAL := 1.0;
    LIM_L : REAL := -1.0E38;
    LIM_H : REAL := 1.0E38;
    RST : BOOL;
  END_VAR
  VAR_OUTPUT
    Y : REAL;
    LIM : BOOL;
  END_VAR
  VAR
    integ : INTEGRATE;
    diff : FT_DERIV;
    YI: REAL;
  END_VAR

  (* run the integrator *)
  IF tn = 0.0 OR rst THEN
    integ(E := FALSE, Y := YI);
    YI := 0.0;
  ELSE
    integ(X := IN, K := 1.0 / TN, E := NOT LIM, Y := YI);
  END_IF;

  (* add up integrator and linear part *)
  Y := KP * (IN + YI);

  (* run differentiator *)
  diff(IN := IN, K := TV);

  (* set lim before differentiator is added to stop integrator if necessary *)
  IF Y > LIM_L AND Y < LIM_H THEN
    LIM := FALSE;
  ELSE
    LIM := TRUE;
  END_IF;

  (* add differential part and limit output Y *)

  Y := LIMIT(LIM_L, Y + KP * diff.out, LIM_H);

(* revision history
  hm 3. jun. 2008   rev 1.0
    original version

  hm  5. nov. 2008  rev 1.1
    changed code to use integrate

  hm  11. mar. 2009 rev 1.2
    real constants updated to new systax using dot
*)
END_FUNCTION_BLOCK

(* @PATH := '\/Engineering\/control' *)
FUNCTION_BLOCK FT_PIW
(*
  FT_PIW is a PI controller.
  The PID controller works according to the fomula Y = IN *(KP+ KI * INTEG(e) ).
  a rst will reset the integrator to 0
  ilim_h and iLim_l set the possible output range of the internal integrator.
  the output flag lim will signal that the output limits are active.
  the controller is equipped with anti wind_up circuitry that stops the integrator when lim_h or lim_l is reached

  default values for KP = 1, KI = 1, ILIM_L = -1E37, iLIM_H = +1E38.
  version 1.0 3. jun 2008
  programmer  hugo
  tested by   tobias
*)
  VAR_INPUT
    IN : REAL;
    KP : REAL := 1.0;
    KI : REAL := 1.0;
    LIM_L : REAL := -1E38;
    LIM_H : REAL := 1E38;
    RST : BOOL;
  END_VAR
  VAR_OUTPUT
    Y : REAL;
    LIM : BOOL;
  END_VAR
  VAR
    integ : FT_INT;
  END_VAR

  (* run integrator *)
  integ(IN := IN, K := KI, RUN := NOT LIM, RST := RST);

  (* set output value *)
  Y := KP * IN + integ.Out;

  (* check for limits and set integrator for anti wind up *)
  IF Y < LIM_L THEN
    Y := LIM_L;
    LIM := TRUE;
  ELSIF Y > LIM_H THEN
    Y := LIM_H;
    LIM := TRUE;
  ELSE
    LIM := FALSE;
  END_IF;

(* revision history
  hm  3. jun. 2008  rev 1.0
    original version
*)
END_FUNCTION_BLOCK

(* @PATH := '\/Engineering\/control' *)
FUNCTION_BLOCK FT_PT2
(*
  FT_PT2 is a 2nd grade filter with programmable times T, D and faktor K.

  version 1.5 11. mar. 2009
  programmer  hugo
  tested by   oscat
*)
  VAR_INPUT
    in : REAL;
    T : TIME;
    D : REAL;
    K : REAL := 1.0;
  END_VAR
  VAR_OUTPUT
    out : REAL;
  END_VAR
  VAR
    init: BOOL;
    int1 : INTEGRATE;
    int2 : INTEGRATE;
    tn: REAL;
    I1, I2 : REAL;
    tn2: REAL;
  END_VAR

  (* startup initialisation *)
  IF NOT init OR T = T#0s THEN
    init := TRUE;
    out := K * in;
    I2 := out;
  ELSE
    TN := TIME_TO_REAL(T) * 1.0E-3;
    tn2 := TN * TN;
    int1(X := in * K / tn2 - I1 * 0.5 * D / TN - I2 / TN2, Y := I1);
    int2(X := I1,Y := I2);
    out := I2;
  END_IF;

(* revision history
  15.1.2007 hm    rev 1.1
    changed formula to new more acurate formula

  hm 15.9.2007    rev 1.2
    deleted unused code for init system time reading tx

  hm  30.11.2007  rev 1.3
    changed out to be K * in during initialization
    avoind divide by 0 if tn = 0

  hm  3. nov. 2008  rev 1.4
    optimized code and fixed a problem with init

  hm  11. mar. 2009 rev 1.5
    real constants updated to new systax using dot
*)
END_FUNCTION_BLOCK

(* @PATH := '\/Engineering\/control' *)
FUNCTION_BLOCK FT_TN16
(*
  FT_TN16 is delay function, it will delay a signal by a specified time : T and will store 16 values of in before they are put thru to out.
  for higher or lower resolution please use FT_TN8 or FT_TN64 instead.

  version 1.1 16 sep 2007
  programmer  hugo
  tested by   tobias
*)
  VAR_INPUT
    in : REAL;
    T : TIME;
  END_VAR
  VAR_OUTPUT
    out : REAL;
    trig : BOOL;
  END_VAR
  VAR
    length : INT := 16;
    X : ARRAY[0..15] OF REAL;
    cnt : INT;
    last : TIME;
    tx: TIME;
    init: BOOL;
  END_VAR

  (* read system time *)
  tx := DWORD_TO_TIME(T_PLC_MS());

  trig := FALSE;
  IF NOT init THEN
    x[cnt] := in;
    init := TRUE;
    last := tx;
  ELSIF tx - last >= T / length THEN
    IF cnt = length - 1 THEN cnt := 0; ELSE cnt := cnt + 1; END_IF;
    Out := X[cnt];
    x[cnt] := in;
    last := tx;
    Trig := TRUE;
  END_IF;

(* revision history
  hm    1. jan 2007 rev 1.0
    original version

  hm    16. sep 2007  rev 1.1
    changes time() to T_plc_ms() for compatibility reasons
*)
END_FUNCTION_BLOCK

(* @PATH := '\/Engineering\/control' *)
FUNCTION_BLOCK FT_TN64
(*
  FT_TN7 is delay function, it will delay a signal by a specified time : T and will store 64 values of in before they are put thru to out.
  if lower resolution is needed, pls use FT_TN8 or FT_TN16 instead.

  version 1.1 15 sep 2007
  programmer  hugo
  tested by   tobias
*)
  VAR_INPUT
    in : REAL;
    T : TIME;
  END_VAR
  VAR_OUTPUT
    out : REAL;
    trig: BOOL;
  END_VAR
  VAR
    length : INT := 64;
    X : ARRAY[0..63] OF REAL;
    cnt : INT;
    last : TIME;
    tx: TIME;
    init: BOOL;
  END_VAR

  (* read system time *)
  tx := DWORD_TO_TIME(T_PLC_MS());

  trig := FALSE;
  IF NOT init THEN
    x[cnt] := in;
    init := TRUE;
    last := tx;
  ELSIF tx - last >= T / length THEN
    IF cnt = length - 1 THEN cnt := 0; ELSE cnt := cnt + 1; END_IF;
    Out := X[cnt];
    x[cnt] := in;
    last := tx;
    trig := TRUE;
  END_IF;

(* revision history
  hm    1. jan 2007   rev 1.0
    original version

  hm    16. sep 2007  rev 1.1
    changes time() to T_plc_ms() for compatibility reasons
*)
END_FUNCTION_BLOCK

(* @PATH := '\/Engineering\/control' *)
FUNCTION_BLOCK FT_TN8
(*
  FT_TN8 is delay function, it will delay a signal by a specified time : T and will store 8 values of in before they are put thru to out.
  if higher resolution is needed, pls use FT_TN16 or FT_TN64 instead.

  version 1.1 15 Sep 2007
  programmer  hugo
  tested by   tobias
*)
  VAR_INPUT
    in : REAL;
    T : TIME;
  END_VAR
  VAR_OUTPUT
    out : REAL;
    trig: BOOL;
  END_VAR
  VAR
    length : INT := 8;
    X : ARRAY[0..7] OF REAL;
    cnt : INT;
    last : TIME;
    tx: TIME;
    init: BOOL;
  END_VAR

  tx := DWORD_TO_TIME(T_PLC_MS());
  trig := FALSE;
  IF NOT init THEN
    x[cnt] := in;
    init := TRUE;
    last := tx;
  ELSIF tx - last >= T / length THEN
    IF cnt = length - 1 THEN cnt := 0; ELSE cnt := cnt + 1; END_IF;
    Out := X[cnt];
    x[cnt] := in;
    last := tx;
    trig := TRUE;
  END_IF;

(* revision history
  hm    1. jan 2007   rev 1.0
    original version

  hm    16. sep 2007  rev 1.1
    changes time() to T_plc_ms() for compatibility reasons
*)
END_FUNCTION_BLOCK

(* @PATH := '\/Engineering\/control' *)
FUNCTION_BLOCK HYST
(*
  This Hystereses function has two modes:
  1. if on > off then Q will be switched high when in > on and switched low when in < off.
  2. if on < off then Q will be switched high when in < on and switched low when in > off.
  the output win will be high when in is between low and high.

  version 1.0 2. jun. 2008
  programmer  hugo
  tested by oscat
*)
  VAR_INPUT
    In : REAL;
    ON : REAL;
    OFF : REAL;
  END_VAR
  VAR_OUTPUT
    Q : BOOL;
    win : BOOL;
  END_VAR

  IF ON >= OFF THEN
    IF IN < OFF THEN
      Q := FALSE;
      WIN := FALSE;
    ELSIF  IN > ON THEN
      Q := TRUE;
      WIN := FALSE;
    ELSE
      WIN := TRUE;
    END_IF;
  ELSE
    IF IN > OFF THEN
      Q := FALSE;
      WIN := FALSE;
    ELSIF  IN < ON THEN
      Q := TRUE;
      WIN := FALSE;
    ELSE
      WIN := TRUE;
    END_IF;
  END_IF;

(* revision history
  hm    2.  jun 2008  rev 1.0
    original version
*)
END_FUNCTION_BLOCK

(* @PATH := '\/Engineering\/control' *)
FUNCTION_BLOCK HYST_1
(*
  this hysteresis function switches the output high if the input signal reaches obove high and will switch to low when the input falls back below low value.
  a separate output mid is set if the input stays between low and high value.

  version 1.1 2. jun. 2008
  programmer  hugo
  tested by oscat
*)
  VAR_INPUT
    In : REAL;
    high : REAL;
    low : REAL;
  END_VAR
  VAR_OUTPUT
    Q : BOOL;
    win : BOOL;
  END_VAR

  IF in < low THEN
    Q := FALSE;
    win := FALSE;
  ELSIF in > high THEN
    Q := TRUE;
    win := FALSE;
  ELSE
    win := TRUE;
  END_IF;

(* revision history
  hm    4.  aug. 2006 rev 1.0
    original version

  hm    2. jun. 2008  rev 1.1
    improved performance
*)
END_FUNCTION_BLOCK

(* @PATH := '\/Engineering\/control' *)
FUNCTION_BLOCK HYST_2
(*
  this hysteresis function switches the output high if the input signal reaches obove val + hys/2 and will switch to low when the input falls back below val - hys/2 value.
  a separate output mid is set if the input stays between low and high value.

  version 1.2 2. jun. 2008
  programmer  oscat
  tested by oscat
*)
  VAR_INPUT
    IN : REAL;
    VAL : REAL;
    HYS : REAL;
  END_VAR
  VAR_OUTPUT
    Q : BOOL;
    WIN: BOOL;
  END_VAR
  VAR
    tmp: REAL;
  END_VAR

  tmp := val - hys * 0.5;
  IF in < tmp THEN
    Q := FALSE;
    win := FALSE;
  ELSIF in > tmp + hys THEN
    Q := TRUE;
    win := FALSE;
  ELSE
    win := TRUE;
  END_IF;

(* revision history
  hm    4. aug 2006 rev 1.0
    original version

  hm    5. jan 2008 rev 1.1
    improved code for better performance

  hm    2. jun. 2008  rev 1.2
    improved performance
*)
END_FUNCTION_BLOCK

(* @PATH := '\/Engineering\/control' *)
FUNCTION_BLOCK HYST_3
(*
  this is a double hysteresis function. Out1 follows a hysteresis function defined by val1and hyst, while out 2 follows val2 and hyst.
  if the input signal is between the two hysteresis switches (val1 and val2) then non of the outputs is active.

  version 1.2 5 jan 2008
  programmer  oscat
  tested by oscat
*)
  VAR_INPUT
    in : REAL;
    hyst : REAL;
    val1 : REAL;
    val2 : REAL;
  END_VAR
  VAR_OUTPUT
    Q1 : BOOL;
    Q2 : BOOL;
  END_VAR
  VAR
    X: REAL;
  END_VAR

  X := hyst * 0.5;
  IF in < val1 - X THEN
    q1 := TRUE;
  ELSIF in > val1 + X THEN
    q1 := FALSE;
  END_IF;
  IF in < val2 - X THEN
    q2 := FALSE;
  ELSIF in > val2 + X THEN
    q2 := TRUE;
  END_IF;

(* revision history
  hm  22. jan 2007  rev 1.0
    original version

  hm  27. dec 2007  rev 1.1
    changed code for better performance

  hm  5. jan 2008 rev 1.2
    further performance iprovements
*)
END_FUNCTION_BLOCK
